(* IEC 61131-3 sources: volt/packages/volt-lsp-iec/test-corpus/lenze-mid/Device/Plc Logic/Application/Library Manager/AlarmManager, 462 files *)

(* ---- ACKNOWLEDGEMETHOD.dut ---- *)
TYPE ACKNOWLEDGEMETHOD :
(
	ACK := 1,
	REP := 2,
	REP_ACK := 3,
	ACK_REP := 6,
	ACK_REP_ACK := 7
);
END_TYPE

(* ---- ALARM_ID.dut ---- *)
TYPE ALARM_ID : UINT;
END_TYPE

(* ---- ALARMBASEPROPERTYINFO.dut ---- *)
TYPE ALARMBASEPROPERTYINFO :
STRUCT
	PVARADR : POINTER TO BYTE;
END_STRUCT
END_TYPE

(* ---- ALARMEVENT.dut ---- *)
TYPE ALARMEVENT :
STRUCT
	USIALARMGROUPID : ALARMGROUP_ID;
	UIALARMID : ALARM_ID;
	LIPUTINTOEVENTQUEUEAT : Timestamp;
END_STRUCT
END_TYPE

(* ---- ALARMGROUP_ID.dut ---- *)
TYPE ALARMGROUP_ID : USINT;
END_TYPE

(* ---- ALARMINDICES.dut ---- *)
TYPE ALARMINDICES :
STRUCT
	M_IALARMGROUPINDEX : INT;
	M_IALARMINDEX : INT;
	M_ICALLERINDEX : INT;
END_STRUCT
END_TYPE

(* ---- ALARMMANAGERCLIENTINFOSTRUCT.dut ---- *)
TYPE ALARMMANAGERCLIENTINFOSTRUCT :
STRUCT
	ITFALARMMANAGERCLIENT : IAlarmManagerClient;
	PARRITFRELEVANTALARMS : POINTER TO ARRAY [0..10] OF IAlarm;
	ICOUNTRELEVANTALARMSLOC : INT;
	DICOUNTRELEVANTALARMSREM : DINT;
	PARRITFACTIVEALARMS : POINTER TO ARRAY [0..10] OF IAlarm;
	ICOUNTACTIVEALARMS : INT;
	PARRITFALARMSFROMHISTORY : POINTER TO ARRAY [0..10] OF IAlarm2;
	PARRALARMSGRPFORHISTORY : POINTER TO ARRAY [0..10] OF POINTER TO AlarmGroupAdapter;
	PARRALARMSCLFORHISTORY : POINTER TO ARRAY [0..10] OF POINTER TO AlarmClassAdapter;
	ICOUNTALARMSFROMHISTORY : INT;
	PARRSTRUCTPROXYREGISTERED : POINTER TO ARRAY [0..10] OF StructProxyRegistered;
	IPROXYCNT : INT;
END_STRUCT
END_TYPE

(* ---- ALARMMANAGERGETALARMSEVENTPARAMS.dut ---- *)
TYPE ALARMMANAGERGETALARMSEVENTPARAMS :
STRUCT
	PSZAPPLNAME : POINTER TO STRING;
	ISKIPROWS : INT;
	IMAXROWS : INT;
	UDICOUNTALARMGROUPS : UDINT;
	PUIARRALARMGROUPS : POINTER TO ARRAY [0..0] OF UDINT;
	UDICOUNTALARMCLASSES : UDINT;
	PUIARRALARMCLASSES : POINTER TO ARRAY [0..0] OF UDINT;
	USIPRIORITYFROM : USINT;
	USIPRIORITYTO : USINT;
	BROWIDVALID : BOOL;
	DIROWID : DINT;
	PBRESULT : POINTER TO BYTE;
	UDIBUFFERSIZE : UDINT;
	UDICOUNTROWS : UDINT;
	UIERROR : UINT;
	BREQUESTHANDLED : BOOL;
END_STRUCT
END_TYPE

(* ---- ALARMMANAGERGETCOUNTEVENTPARAMS.dut ---- *)
TYPE ALARMMANAGERGETCOUNTEVENTPARAMS :
STRUCT
	PSZAPPLNAME : POINTER TO STRING;
	UDICOUNTALARMGROUPS : UDINT;
	PUIARRALARMGROUPS : POINTER TO ARRAY [0..0] OF UDINT;
	UDICOUNTALARMCLASSES : UDINT;
	PUIARRALARMCLASSES : POINTER TO ARRAY [0..0] OF UDINT;
	USIPRIORITYFROM : USINT;
	USIPRIORITYTO : USINT;
	UDICOUNT : UDINT;
	BREQUESTHANDLED : BOOL;
END_STRUCT
END_TYPE

(* ---- ALARMRECORD.dut ---- *)
TYPE ALARMRECORD :
STRUCT
	IRECORDID : INT := -1;
	UICLIENT : UINT;
	IALARMGROUP : INT;
	PAITFALARMGROUP : POINTER TO ARRAY [0..9] OF IAlarmGroup;
	IALARMCLASS : INT;
	PAITFALARMCLASS : POINTER TO ARRAY [0..9] OF IAlarmClass;
	IALARMCLASSINSERT : INT;
END_STRUCT
END_TYPE

(* ---- ALARMSTATE.dut ---- *)
TYPE ALARMSTATE :
(
	NOTDEFINED := 16#FF,
	NORMAL := 0,
	ACTIVE := 2,
	WAITINGFORCONFIRMATION := 3,
	ACTIVEACKNOWLEDGED := 4,
	INACTIVEUNACKNOWLEDGED := 5,
	PENDING := 1
);
END_TYPE

(* ---- ALARMSTATETRANSITION.dut ---- *)
TYPE ALARMSTATETRANSITION :
(
	NOTRANSITION := 0,
	PENDING := -1,
	ACTIVATE := 1,
	DEACTIVATE := 2,
	ACKNOWLEDGE := 3,
	CONFIRM := 4,
	REALARM := 5
);
END_TYPE

(* ---- ALARMSTORAGELATCHVARIABLE.dut ---- *)
TYPE ALARMSTORAGELATCHVARIABLE :
STRUCT
	M_BYTYPE : BYTE;
	M_LIVALUE : LINT;
	M_XVALUENULL : BOOL;
END_STRUCT
END_TYPE

(* ---- ALARMSTORAGESTATICDATA.dut ---- *)
TYPE ALARMSTORAGESTATICDATA :
STRUCT
	LITIMESTAPLAST : TIMESTAMP;
	LITIMESTAPACTIVE : TIMESTAMP;
	LITIMESTAPINACTIVE : TIMESTAMP;
	LITIMESTAPACKNOWLEDGE : TIMESTAMP;
	IOFFSETLAST : INT := -1;
	IOFFSETACTIVE : INT := -1;
	IOFFSETINACTIVE : INT := -1;
	IOFFSETACKNOWLEDGE : INT := -1;
	LITRIGGERVALUEVAL : LINT;
	ITRIGGERVALUETYPE : TypeClass;
	UDIALARMID : UDINT;
	UDIALARMGROUPID : UDINT;
	UDIALARMCLASSID : UDINT;
	ESTATE : AlarmState;
	USIPRIORITY : USINT;
	LIREMOTEDEVICEVAL : LINT;
	PWSCMTACTIVEACK : POINTER TO WSTRING;
	PWSCMTNORMAL : POINTER TO WSTRING;
	PWSCMTACTIVE : POINTER TO WSTRING;
	PWSCMTWAITINGCONF : POINTER TO WSTRING;
	PWSUSERIDACTIVEACK : POINTER TO WSTRING;
	PWSUSERIDNORMAL : POINTER TO WSTRING;
	PWSUSERIDACTIVE : POINTER TO WSTRING;
	PWSUSERIDWAITINGCONF : POINTER TO WSTRING;
	IDROW : CAA.IDENT;
END_STRUCT
END_TYPE

(* ---- ALARMSTRUCTFONT.dut ---- *)
TYPE ALARMSTRUCTFONT :
STRUCT
	SNAME : STRING := 'Arial';
	IHEIGHT : INT := 12;
	DWFLAGS : DWORD := 16#0;
	DWCHARSET : DWORD := 16#0;
	DWCOLOR : DWORD := 16#0;
END_STRUCT
END_TYPE

(* ---- ALARMUNIONBYTEORDERTEST.dut ---- *)
TYPE ALARMUNIONBYTEORDERTEST :
UNION
	W : WORD;
	BTS : ARRAY [0..1] OF BYTE;
END_UNION
END_TYPE

(* ---- CONFIGURABLEEXPRESSION.dut ---- *)
TYPE CONFIGURABLEEXPRESSION :
(
	OBSERVEDEXPRESSION := 0,
	LATCHVAR1 := 1,
	LATCHVAR2 := 2,
	LASTLATCHVARIABLE := 1000
);
END_TYPE

(* ---- DISPLAYOPTIONS.dut ---- *)
TYPE DISPLAYOPTIONS :
STRUCT
	FONT : AlarmStructFont;
	DWBACKGROUNDCOLOR : DWORD := 16#FFFFFF;
	SBITMAPID : STRING;
	XTRANSPARENT : BOOL;
	DWTRANSPARENTCOLOR : DWORD;
END_STRUCT
END_TYPE

(* ---- EALARMBYTEORDER.dut ---- *)
TYPE EALARMBYTEORDER :
(
	INTEL,
	MOTOROLA,
	UNKNOWN
);
END_TYPE

(* ---- EALARMCOMMENT.dut ---- *)
TYPE EALARMCOMMENT :
(
	NO_COMMENT,
	COMMENT_NORMAL,
	COMMENT_ACTIVE_ACK
);
END_TYPE

(* ---- EALARMCOMPARABLE.dut ---- *)
TYPE EALARMCOMPARABLE :
(
	FIRST_ENTRY := 0,
	TIMESTAMP_LAST := 0,
	TIMESTAMP_ACTIVE := 1,
	TIMESTAMP_INACTIVE := 2,
	TIMESTAMP_ACKNOWLEDGE := 3,
	VALUE := 4,
	MESSAGE := 5,
	PRIORITY := 6,
	ALARM_CLASS := 7,
	STATE := 8,
	REM_DEVICE := 9,
	COMMENT_ACK := 10,
	USERID_ACK := 11,
	LAST_ENTRY := 11
);
END_TYPE

(* ---- EALARMSTORAGEMIRRORSTATE.dut ---- *)
TYPE EALARMSTORAGEMIRRORSTATE :
(
	NOTYETMIRRORED,
	MIRRORINGSTARTED,
	ADDITIONALREADCALLREQUIRED,
	COMPLETELYMIRRORED,
	ERROR,
	RELOADREQUIRED
);
END_TYPE

(* ---- EALARMSTORAGEOBJECT.dut ---- *)
TYPE EALARMSTORAGEOBJECT :
(
	IX_MIN := 0,
	TBL_ALARM := IX_MIN,
	TBL_METADATA := 1,
	TBL_VERSION := 2,
	IDX_TSLAST := 3,
	IDX_GROUP_TSLAST := 4,
	IDX_CLASS_TSLAST := 5,
	TBL_LATCH_VAR_STRINGS := 6,
	IDX_LATCH_VAR_STRINGS := 7,
	IDX_LATCH1_TSLAST := 8,
	IX_LAST := IDX_LATCH1_TSLAST
);
END_TYPE

(* ---- EALARMSTORAGEREADERERRORS.dut ---- *)
TYPE EALARMSTORAGEREADERERRORS :
(
	NOERROR := CmpErrors.Errors.ERR_OK,
	WRONGPARAMETER := CmpErrors.Errors.ERR_PARAMETER,
	NOMEMORY := CmpErrors.Errors.ERR_NOMEMORY,
	NOOBJECT := CmpErrors.Errors.ERR_NO_OBJECT,
	ADDITIONALREADCALLREQUIRED := CmpErrors.Errors.ERR_PENDING,
	INVALIDCALL := 20002
);
END_TYPE

(* ---- EALARMTYPE.dut ---- *)
TYPE EALARMTYPE :
(
	UNDEFINED := 0,
	ALARM := 1,
	EVENT := 2,
	IMPLICITLYACKNOWLEDGEDEVENT := 3,
	ALARMAPI := 4
);
END_TYPE

(* ---- ECOMPARABLETYPE.dut ---- *)
TYPE ECOMPARABLETYPE :
(
	TYPE_UNDEFINED := 0,
	TYPE_BOOL := 1,
	TYPE_NUMERIC := 2,
	TYPE_STRING := 3
);
END_TYPE

(* ---- EDBACTIVEINDEX.dut ---- *)
TYPE EDBACTIVEINDEX :
(
	NOT_DEFINED := 0,
	TIMESTAMP,
	GROUP,
	EDB_CLASS,
	LATCH1
);
END_TYPE

(* ---- EDBTYPE.dut ---- *)
TYPE EDBTYPE :
(
	NOT_DEFINED := 0,
	SQL,
	MEMORY
);
END_TYPE

(* ---- EFILTERLATCHCONTENT.dut ---- *)
TYPE EFILTERLATCHCONTENT :
(
	NOT_SET := -1,
	DISABLE := 0,
	STR := 1,
	IEC := 2,
	NUMBER := 3
);
END_TYPE

(* ---- EFILTERTIMERANGETYPE.dut ---- *)
TYPE EFILTERTIMERANGETYPE :
(
	NOT_SET := -1,
	DISABLE := 0,
	ENABLE := 1
);
END_TYPE

(* ---- ELOCALBUFFERCURSORSTATE.dut ---- *)
TYPE ELOCALBUFFERCURSORSTATE :
(
	EOF := -3,
	CLOSED := -2,
	OPEN := -1
);
END_TYPE

(* ---- ENUMERICCOMPARISON.dut ---- *)
TYPE ENUMERICCOMPARISON :
(
	AS_LINT := 0,
	AS_REAL := 1,
	AS_LREAL := 2
);
END_TYPE

(* ---- EVTPARAM_CHANNELCLOSED.dut ---- *)
TYPE EVTPARAM_CHANNELCLOSED :
STRUCT
	UICLIENT : UINT;
	UICHANNELHANDLE : UINT;
	ERRREASON : RTS_IEC_RESULT;
END_STRUCT
END_TYPE

(* ---- FILELIMIT.dut ---- *)
TYPE FILELIMIT :
(
	NOLIMIT := 0,
	RECORDS := 1,
	SIZE := 2
);
END_TYPE

(* ---- HISTORICALACTIVEALARMROWID.dut ---- *)
TYPE HISTORICALACTIVEALARMROWID :
STRUCT
	DWROWID : DWORD;
	LITS : LINT;
END_STRUCT
END_TYPE

(* ---- LATCHVARIABLE.dut ---- *)
TYPE LATCHVARIABLE :
STRUCT
	M_BYTYPE : BYTE;
	M_LIVALUE : LINT;
END_STRUCT
END_TYPE

(* ---- LOCALBUFFERDATABASEACCESSCONTEXT.dut ---- *)
TYPE LOCALBUFFERDATABASEACCESSCONTEXT :
STRUCT
	M_HSEMTRANSACTION : RTS_IEC_HANDLE := RTS_INVALID_HANDLE;
	M_DICURSORINDEX : DINT := ELocalBufferCursorState.Closed;
	M_PALICURRALARM : POINTER TO ARRAY [0..0] OF LINT;
	M_CBPSTRINGLATCHVARIABLE : CharBufferPtr;
	M_XISONLYONEALARMGROUPSELECTED : BOOL;
	M_XISONLYONEALARMCLASSSELECTED : BOOL;
	M_ELASTERROR : STO.ERROR;
END_STRUCT
END_TYPE

(* ---- MONITORDBSTATUS.dut ---- *)
TYPE MONITORDBSTATUS :
STRUCT
	DBTYPE : EDBType;
	ACTIVEINDEX : EDBActiveIndex;
	IERROR : INT;
	SFUNCTION : STRING;
	IACTION : INT;
END_STRUCT
END_TYPE

(* ---- MONITORFILTERBYDATETIME.dut ---- *)
TYPE MONITORFILTERBYDATETIME :
STRUCT
	FILTERTARGET : EFilterTimeRangeType;
	DTFROMVALUE : DATE_AND_TIME;
	DTTOVALUE : DATE_AND_TIME;
END_STRUCT
END_TYPE

(* ---- MONITORFILTERBYLATCH.dut ---- *)
TYPE MONITORFILTERBYLATCH :
STRUCT
	FILTERLATCHCONTENT : EFilterLatchContent;
	VTYPE : Visu_Types;
	LIVALUE : LINT;
	RVALUE : REAL;
	LRVALUE : LREAL;
	WSSTRVALUE : WSTRING(255);
END_STRUCT
END_TYPE

(* ---- PLACEHOLDERANALYZATIONSTATE.dut ---- *)
TYPE PLACEHOLDERANALYZATIONSTATE :
(
	NOTAVAILABLE := 16#0,
	TOOMANYPLACEHOLDERS := 16#1,
	INVALIDPLACEHOLDER := 16#2,
	CYCLICALLYREPAINTREQUIRED := 16#4,
	DONE := 16#10
);
END_TYPE

(* ---- PLACEHOLDERDESCRIPTION.dut ---- *)
TYPE PLACEHOLDERDESCRIPTION :
STRUCT
	M_EPLACEHOLDER : Placeholder;
	M_PCBSPLACEHOLDER : POINTER TO CharBufferString;
	M_XSUPPORTSFORMATSTRING : BOOL;
	M_XINHIBITSOPTIMIZATION : BOOL;
	M_XREQUIREDCYCLICALLYREPAINT : BOOL;
	M_XINHIBITMULTIPLEUSAGE : BOOL;
	M_PCBSRELATEDPLACEHOLDERSUBSTRING : POINTER TO CharBufferString;
	M_PCBSRELATEDPLACEHOLDERBRACKET : POINTER TO CharBufferString;
END_STRUCT
END_TYPE

(* ---- PLACEHOLDERINFO.dut ---- *)
TYPE PLACEHOLDERINFO :
STRUCT
	M_APLACEHOLDEROCCURRENCE : ARRAY [0..(AlarmConstants.COUNT_PLACEHOLDER - 1)] OF PlaceholderOccurrence;
	M_SICOUNTPLACEHOLDERS : SINT := -1;
	M_EPLACEHOLDERANALYZATIONSTATE : PlaceholderAnalyzationState;
END_STRUCT
END_TYPE

(* ---- PLACEHOLDERSCANNERSTATE.dut ---- *)
TYPE PLACEHOLDERSCANNERSTATE :
(
	START := 0,
	SKIPWHITESPACE := 1,
	SCANFORMAT := 2,
	END := 3,
	ERROR := 255
);
END_TYPE

(* ---- PROXYENUMSTATE.dut ---- *)
TYPE PROXYENUMSTATE :
(
	NOTRUNNING,
	PREPARATION,
	CHECKDATA,
	RUN
);
END_TYPE

(* ---- PROXYSTRUCTALARM.dut ---- *)
TYPE PROXYSTRUCTALARM :
STRUCT
	UIALARMID : ALARM_ID;
	UDIALARMINTERNALID : UDINT;
	UDIALARMGROUPINTERNALID : UDINT;
	UDIALARMCLASSINTERNALID : UDINT;
	SALARMID : STRING;
	XACK : BOOL;
END_STRUCT
END_TYPE

(* ---- PROXYSTRUCTALARMCLASS.dut ---- *)
TYPE PROXYSTRUCTALARMCLASS :
STRUCT
	UDIINTERNALID : UDINT;
	SNAME : STRING;
	USIPRIORITY : USINT;
	XACKNOWLEDGESEPARATELY : BOOL;
	ADISPLAYOPTIONS : ARRAY [AlarmState.Normal..AlarmState.ActiveAcknowledged] OF DisplayOptions;
	AXDISPLAYOPTIONSSET : ARRAY [AlarmState.Normal..AlarmState.ActiveAcknowledged] OF BOOL;
END_STRUCT
END_TYPE

(* ---- PROXYSTRUCTALARMCLASSDESC.dut ---- *)
TYPE PROXYSTRUCTALARMCLASSDESC :
STRUCT
	XVALID : BOOL;
	SNAME : STRING;
	USIPRIORITY : USINT;
	UDIINTERNALID : UDINT;
END_STRUCT
END_TYPE

(* ---- PROXYSTRUCTALARMDESC.dut ---- *)
TYPE PROXYSTRUCTALARMDESC :
STRUCT
	XVALID : BOOL;
	SALARMID : STRING;
	UIALARMID : ALARM_ID;
	UDIALARMINTERNALID : UDINT;
	UDIALARMGROUPINTERNALID : UDINT;
END_STRUCT
END_TYPE

(* ---- PROXYSTRUCTALARMGROUP.dut ---- *)
TYPE PROXYSTRUCTALARMGROUP :
STRUCT
	UDIINTERNALID : UDINT;
	SNAME : STRING;
	STEXTLIST : STRING;
END_STRUCT
END_TYPE

(* ---- PROXYSTRUCTALARMGROUPDESC.dut ---- *)
TYPE PROXYSTRUCTALARMGROUPDESC :
STRUCT
	XVALID : BOOL;
	SNAME : STRING;
	STEXTLIST : STRING;
	UDIINTERNALID : UDINT;
END_STRUCT
END_TYPE

(* ---- PROXYSTRUCTCLASSREMAP.dut ---- *)
TYPE PROXYSTRUCTCLASSREMAP :
STRUCT
	SCLASSORIGINAL : STRING;
	SCLASSNEW : STRING;
END_STRUCT
END_TYPE

(* ---- PROXYSTRUCTDSCHANNELPARAM.dut ---- *)
TYPE PROXYSTRUCTDSCHANNELPARAM :
STRUCT
	ITFDATASOURCESMGR : IDatasources.IDatasourcesMgr;
	PSDSNAME : POINTER TO STRING;
	ILATCHVARSNUM : INT;
	PSALMSTATETRANSCOUNTER : POINTER TO STRING;
	PALMSTATETRANSCOUNTER : __XWORD;
	TYPEALMSTATETRANSCOUNTER : TypeClass;
	PSALMSTORAGECOUNTER : POINTER TO STRING;
	PALMSTORAGECOUNTER : __XWORD;
	TYPEALMSTORAGECOUNTER : TypeClass;
END_STRUCT
END_TYPE

(* ---- PROXYSTRUCTERROR.dut ---- *)
TYPE PROXYSTRUCTERROR :
STRUCT
	UDIERROR : UDINT;
	LTTIMESTAMP : LTIME;
	SMSG : STRING(20);
END_STRUCT
END_TYPE

(* ---- PROXYSTRUCTHISTORICALALARMACTIVE.dut ---- *)
TYPE PROXYSTRUCTHISTORICALALARMACTIVE :
STRUCT
	DWROWIDLOCAL : DWORD := AlarmConstants.INVALID_ROWID;
	DWROWIDREMOTE : DWORD := AlarmConstants.INVALID_ROWID;
	LITSACTIVEREMOTE : LINT;
	ESTATELAST : AlarmState := AlarmState.NotDefined;
END_STRUCT
END_TYPE

(* ---- PROXYSTRUCTINITIALIZE.dut ---- *)
TYPE PROXYSTRUCTINITIALIZE :
STRUCT
	PSPROXYNAME : POINTER TO STRING;
	ITFPROXYCOMMCHANNEL : IProxyCommChannel;
	PSAPPNAME : POINTER TO STRING;
	PAALARMGROUPS : POINTER TO ARRAY [0..9] OF STRING;
	IALARMGROUPSNUM : INT;
	PACLASSREMAP : POINTER TO ARRAY [0..9] OF ProxyStructClassReMap;
	ICLASSREMAPNUM : INT;
END_STRUCT
END_TYPE

(* ---- PROXYSTRUCTMONITOR.dut ---- *)
TYPE PROXYSTRUCTMONITOR :
STRUCT
	SNAME : STRING;
	ESTATE : ProxyEnumState;
	IALARMCLASSNUM : INT;
	IALARMGROUPSNUM : INT;
	DIALARMNUM : DINT;
	ILATCHVARSNUM : INT;
	IACTIVEALARMS : INT;
	DIHISTACTIVEALMSCNT : DINT;
	IHISTROWALMSCNT : INT;
	IHISTROWACTIVEALMSCNT : INT;
	XHASSTORAGE : BOOL;
	DWROWIDFIRSTREMDB : DWORD;
	DWROWIDLASTREMDB : DWORD;
	DWROWIDLASTLOCDB : DWORD;
	DIWRITEDBCNTTOT : DINT;
	IWRITEDBCNT : INT;
	TWRITEDBDURATIONLAST : TIME;
	DITOTMEM : DINT;
	DIHISTACTIVEALMSSIZE : DINT;
	IHISTROWALMSSIZE : INT;
	IHISTROWACTIVEALMSSIZE : INT;
	LIBVERALMMAN : VERSION;
END_STRUCT
END_TYPE

(* ---- PROXYSTRUCTMONITORALARMCLASSDESC.dut ---- *)
TYPE PROXYSTRUCTMONITORALARMCLASSDESC :
STRUCT
	SNAME : STRING;
	UDIINTERNALID : UDINT;
	USIPRIORITY : USINT;
	XACKNOWLEDGESEPARATELY : BOOL;
END_STRUCT
END_TYPE

(* ---- PROXYSTRUCTMONITORALARMDESC.dut ---- *)
TYPE PROXYSTRUCTMONITORALARMDESC :
STRUCT
	SALARMID : STRING;
	UIALARMID : ALARM_ID;
	UDIALARMINTERNALID : UDINT;
	UDIALARMGROUPINTERNALID : UDINT;
	UDIALARMCLASSINTERNALID : UDINT;
END_STRUCT
END_TYPE

(* ---- PROXYSTRUCTMONITORALARMGROUPDESC.dut ---- *)
TYPE PROXYSTRUCTMONITORALARMGROUPDESC :
STRUCT
	SNAME : STRING;
	UDIINTERNALID : UDINT;
	STEXTLIST : STRING;
END_STRUCT
END_TYPE

(* ---- PROXYSTRUCTMONITORREQUEST.dut ---- *)
TYPE PROXYSTRUCTMONITORREQUEST :
STRUCT
	ITASKID : INT := ProxyConstants.REQ_ID_NONE;
	AFIFOERRORS : ARRAY [1..ProxyConstants.FIFO_ERROR_SIZE] OF ProxyStructError;
	UDIERRCOUNT : UDINT;
	LTELAPTIME : LTIME;
	TREQDURATIONLAST : TIME;
	TREQDURATIONAVG : TIME;
	TREQDURATIONMIN : TIME;
	TREQDURATIONMAX : TIME;
	UDIREQDURATIONBUILDREQ : UDINT;
	UDIREQDURATIONWAITANS : UDINT;
	UDIREQDURATIONELABANS : UDINT;
	UDIREQCOUNT : UDINT;
	UDIREQCOUNTCLOSED : UDINT;
END_STRUCT
END_TYPE

(* ---- PROXYSTRUCTPARAM.dut ---- *)
TYPE PROXYSTRUCTPARAM :
STRUCT
	DWBASETIME : DWORD;
	DWACTALMTIME : DWORD;
	DWHISALMTIME : DWORD;
	DWACKALMTIME : DWORD;
	TTIMEOUT : TIME := TIME#5s0ms;
END_STRUCT
END_TYPE

(* ---- PROXYSTRUCTRECORD.dut ---- *)
TYPE PROXYSTRUCTRECORD :
STRUCT
	IRECORDID : INT;
	IALARMCLASSNUM : INT;
	DIALARMNUM : DINT;
	ILATCHVARSNUM : INT;
	PAALARMGROUPS : POINTER TO ARRAY [0..9] OF STRING;
	IALARMGROUPSNUM : INT;
	PACLASSREMAP : POINTER TO ARRAY [0..9] OF ProxyStructClassReMap;
	ICLASSREMAPNUM : INT;
	PAACTIVEALARMOBJSTUBS : POINTER TO ARRAY [0..100] OF POINTER TO ProxyFbAlarmMetaObjectStub;
	DIALMOBJSTUBSALLOC : DINT;
	PAACTIVEALARMCONTAINER : POINTER TO ARRAY [0..100] OF POINTER TO AlarmContainer;
	DIALMCONTAINERALLOC : DINT;
	DIACTIVEALARMS : DINT;
	PASTRUCTALARMDESCRIPTION : POINTER TO ARRAY [0..100] OF POINTER TO ProxyStructAlarm;
	DIALARMDESCALLOC : DINT;
	PASTRUCTALARMGROUPDESCRIPTION : POINTER TO ARRAY [0..100] OF POINTER TO ProxyStructAlarmGroup;
	IALARMGROUPDESCALLOC : INT;
	PASTRUCTALARMCLASSDESCRIPTION : POINTER TO ARRAY [0..100] OF POINTER TO ProxyStructAlarmClass;
	IALARMCLASSDESCALLOC : INT;
END_STRUCT
END_TYPE

(* ---- PROXYSTRUCTTASKCALL.dut ---- *)
TYPE PROXYSTRUCTTASKCALL :
STRUCT
	ITASKID : INT;
	DWSCHEDUL : DWORD;
	TTIMEOUT : TIME;
	XDONEOK : BOOL;
	XLOCK : BOOL;
	HLOCK : RTS_IEC_HANDLE;
	DWSCHEDULCNT : DWORD;
END_STRUCT
END_TYPE

(* ---- SCALARTYPE.dut ---- *)
TYPE SCALARTYPE :
UNION
	COMPBYTE : BYTE;
	COMPWORD : WORD;
	COMPDWORD : DWORD;
	COMPLWORD : LWORD;
	COMPSINT : SINT;
	COMPUSINT : USINT;
	COMPINT : INT;
	COMPUINT : UINT;
	COMPDINT : DINT;
	COMPUDINT : UDINT;
	COMPLINT : LINT;
	COMPULINT : ULINT;
	COMPBOOL : BOOL;
	COMPREAL : REAL;
	COMPLREAL : LREAL;
END_UNION
END_TYPE

(* ---- SQLITEDATABASEACCESSCONTEXT.dut ---- *)
TYPE SQLITEDATABASEACCESSCONTEXT :
STRUCT
	M_ITFTABLELATCHVARVALUES : STO.ITable;
	M_ITFCURSORLATCHVARVALUES : STO.ICursor;
	M_ITFROWLATCHVARVALUES : STO.IRow;
	M_IDTBLLATCHVARSTRINGS : CAA.IDENT;
	M_IDIDXLATCHVARSTRINGS : CAA.IDENT;
	M_ITFTRANSACTION : STO.ITransaction;
	M_ITFTABLE : STO.ITable;
	M_ITFCURSOR : STO.ICursor;
	M_ITFROW : STO.IRow;
	M_IDINDEX : CAA.IDENT;
	M_EINDEX : EAlarmStorageObject;
	M_ELASTERROR : STO.ERROR;
END_STRUCT
END_TYPE

(* ---- STORAGETASKINFO.dut ---- *)
TYPE STORAGETASKINFO :
STRUCT
	XTASKACTIVE : BOOL;
	PTASKINFO : POINTER TO CmpIecTask.Task_Info2;
END_STRUCT
END_TYPE

(* ---- STRINGCONTAINERBUFFERINFO.dut ---- *)
TYPE STRINGCONTAINERBUFFERINFO :
STRUCT
	PUDIBUFFERSIZE : POINTER TO UDINT;
	PUDIFIRSTFREEPOSITION : POINTER TO UDINT;
	PBYFIRSTPOSITION : POINTER TO BYTE;
	PBYFIRSTFREEPOSITION : POINTER TO BYTE;
END_STRUCT
END_TYPE

(* ---- STRUCTPROXYREGISTERED.dut ---- *)
TYPE STRUCTPROXYREGISTERED :
STRUCT
	ITFPROXY : IProxy;
	DIALM : DINT;
END_STRUCT
END_TYPE

(* ---- STRUFILTERREMOTEALM.dut ---- *)
TYPE STRUFILTERREMOTEALM :
STRUCT
	SPROXYNAME : STRING;
	DIID : DINT;
END_STRUCT
END_TYPE

(* ---- SWAPHELPER_UNION.dut ---- *)
TYPE SWAPHELPER_UNION :
UNION
	COMPBYTE : BYTE;
	COMPWORD : WORD;
	COMPDWORD : DWORD;
	COMPLWORD : LWORD;
END_UNION
END_TYPE

(* ---- TIMESTAMP.dut ---- *)
TYPE TIMESTAMP : LINT;
END_TYPE

(* ---- ALARMCONSTANTS.gvl ---- *)
VAR_GLOBAL
	NULL : POINTER TO BYTE := 0;
	MAX_PLACEHOLDER_LENGTH : BYTE := 25;
	MAX_PLACEHOLDER_REPLACEMENT_LENGTH : WORD := 255;
	REPL_AMP_ANSI : DWORD := 16#0;
	REPL_AMP_UNICODE : DWORD := 16#1;
	ALARM_MESSAGEBUFFER_SIZE : WORD := 500;
	MAX_MESSAGE_SIZE : WORD := 256;
	ALARM_SEPARATOR : STRING(1) := '$T';
	ALARMGROUP_SEPARATOR : STRING(1) := '|';
	SLEEP_TIME : UDINT := 5;
	RETRY_COUNT : INT := 10;
	NOT_RELEVANT : ALARM_ID := 65535;
	TICKS_1_1_1970 : ULINT := 116444736000000000;
	DIVISOR_TO_SECONDS : LINT := ((1000 * 1000) * 10);
	FMT_INT : BYTE := 0;
	FMT_LONG : BYTE := 1;
	FMT_FLOAT : BYTE := 2;
	FMT_STRING : BYTE := 3;
	FMT_WSTRING : BYTE := 4;
	FMT_FIRST_FORMAT_STRING : BYTE := FMT_INT;
	FMT_LAST_FORMAT_STRING : BYTE := FMT_WSTRING;
	PLH_FIRST_PLACEHOLDER : Placeholder := Placeholder.PLH_ALARM;
	PLH_LAST_PLACEHOLDER : Placeholder := Placeholder.PLH_TRIGGERVALUE;
	COUNT_PLACEHOLDER : BYTE := 22;
	INVALID_ROWID : CAA.IDENT := 0;
	LESS : INT := -1;
	EQUAL : INT := 0;
	GREATER : INT := 1;
	RECORD_ID_TEST : INT := 16#7FFF;
	RECORD_ID_TEST2 : INT := 16#7FFE;
	MAX_LATCH_VARS : INT := 10;
	SIZE_HIST_ACTIVE_ALM : INT := 250;
	VISU_TYPES_TYPE_LDATE : INT := 33;
	VISU_TYPES_TYPE_LDT : INT := 34;
	VISU_TYPES_TYPE_LTOD : INT := 35;
	ALARM_STORAGE_TASK_NAME : STRING := 'Visu_AlarmStorageTask';
END_VAR

(* ---- ALARMGLOBALS.gvl ---- *)
VAR_GLOBAL
	G_ACK_ALARMSTATEMACHINE : Ack_AlarmStateMachine;
	G_ACK_REP_ALARMSTATEMACHINE : Ack_Rep_AlarmStateMachine;
	G_ACK_REP_ACK_ALARMSTATEMACHINE : Ack_Rep_Ack_AlarmStateMachine;
	G_REP_ACK_ALARMSTATEMACHINE : Rep_Ack_AlarmStateMachine;
	G_REP_ALARMSTATEMACHINE : Rep_AlarmStateMachine;
	G_ACK_ALARMSTATEMACHINE_NOCONFIRM : Ack_AlarmStateMachine_NoConfirm;
	G_ACK_REP_ALARMSTATEMACHINE_NOCONFIRM : Ack_Rep_AlarmStateMachine_NoConfirm;
	G_ACK_REP_ACK_ALARMSTATEMACHINE_NOCONFIRM : Ack_Rep_Ack_AlarmStateMachine_NoConfirm;
	G_REP_ACK_ALARMSTATEMACHINE_NOCONFIRM : Rep_Ack_AlarmStateMachine_NoConfirm;
	G_ALARMHANDLER_INST : StandardAlarmHandler;
	G_ALARMHANDLER : IAlarmHandler9 := g_AlarmHandler_Inst;
	G_ALARMHANDLERBASE : IAlarmHandlerBase := g_AlarmHandler_Inst;
	G_ALARMHANDLERREMOTE : IAlarmHandlerRemote := g_AlarmHandler_Inst;
	G_ALARMHANDLERREMOTEMONITOR : IAlarmHandlerRemoteMonitor := g_AlarmHandler_Inst;
	G_ALARMSTORAGEQUEUE : AlarmStorageQueue;
	G_DIALARMSTATETRANSITIONCOUNTER : DINT;
	G_DIALARMSTORAGECOUNTER : DINT;
	STATE : INT;
	G_STAPPLICATIONNAME : STRING;
	G_PAPPLICATION : POINTER TO CmpApp.APPLICATION := RTS_INVALID_HANDLE;
	G_ERRORHANDLER : DatabaseAccessErrorHandler;
	G_BBYTEORDERDETERMINED : BOOL := FALSE;
	G_XMETADATAFILECREATED : BOOL := FALSE;
	G_SDATEFORMAT : STRING := 'dd.MM.yyyy';
	G_STIMEFORMAT : STRING := 'HH:mm:ss';
	G_DATEFORMATTER : STU.DateFormatter;
	G_TIMEFORMATTER : STU.TimeFormatter;
	G_TYPEDVALUEFORMATTER : TypedValueFormatter;
	G_SALARMSTATETEXTLISTNAME : STRING := 'AlarmManager.TL_AlarmStatus';
	COMPONENT_NAME : STRING := 'AlarmManager';
	G_STRINGPLACEHOLDERDATE : CharBufferString;
	G_STRINGPLACEHOLDERDATE2 : CharBufferString;
	G_STRINGPLACEHOLDERALLDEFAULT : CharBufferString;
	G_STRINGPLACEHOLDERMESSAGE : CharBufferString;
	G_STRINGPLACEHOLDERTIME : CharBufferString;
	G_STRINGPLACEHOLDERTIME2 : CharBufferString;
	G_STRINGPLACEHOLDERSTATE : CharBufferString;
	G_STRINGPLACEHOLDERSTATE2 : CharBufferString;
	G_STRINGPLACEHOLDEREXPRESSION : CharBufferString;
	G_STRINGPLACEHOLDEREXPRESSION2 : CharBufferString;
	G_STRINGPLACEHOLDERPRIORITY : CharBufferString;
	G_STRINGPLACEHOLDERPRIORITY2 : CharBufferString;
	G_STRINGPLACEHOLDERCLASS : CharBufferString;
	G_STRINGPLACEHOLDERCLASS2 : CharBufferString;
	G_STRINGPLACEHOLDERALARMID : CharBufferString;
	G_STRINGPLACEHOLDERCURRENTVALUE : CharBufferString;
	G_STRINGPLACEHOLDERCURRENTVALUE2 : CharBufferString;
	G_STRINGPLACEHOLDERTRIGGERVALUE : CharBufferString;
	G_STRINGPLACEHOLDERTRIGGERVALUE2 : CharBufferString;
	G_STRINGPLACEHOLDERLATCH : CharBufferString;
	G_STRINGPLACEHOLDERLATCHWITHOPENINGBRACKET : CharBufferString;
	G_STRINGPLACEHOLDERALARM : CharBufferString;
	G_WSTRINGPLACEHOLDERDATE : CharBufferString;
	G_WSTRINGPLACEHOLDERDATE2 : CharBufferString;
	G_WSTRINGPLACEHOLDERALLDEFAULT : CharBufferString;
	G_WSTRINGPLACEHOLDERMESSAGE : CharBufferString;
	G_WSTRINGPLACEHOLDERTIME : CharBufferString;
	G_WSTRINGPLACEHOLDERTIME2 : CharBufferString;
	G_WSTRINGPLACEHOLDERSTATE : CharBufferString;
	G_WSTRINGPLACEHOLDERSTATE2 : CharBufferString;
	G_WSTRINGPLACEHOLDEREXPRESSION : CharBufferString;
	G_WSTRINGPLACEHOLDEREXPRESSION2 : CharBufferString;
	G_WSTRINGPLACEHOLDERPRIORITY : CharBufferString;
	G_WSTRINGPLACEHOLDERPRIORITY2 : CharBufferString;
	G_WSTRINGPLACEHOLDERCLASS : CharBufferString;
	G_WSTRINGPLACEHOLDERCLASS2 : CharBufferString;
	G_WSTRINGPLACEHOLDERALARMID : CharBufferString;
	G_WSTRINGPLACEHOLDERCURRENTVALUE : CharBufferString;
	G_WSTRINGPLACEHOLDERCURRENTVALUE2 : CharBufferString;
	G_WSTRINGPLACEHOLDERTRIGGERVALUE : CharBufferString;
	G_WSTRINGPLACEHOLDERTRIGGERVALUE2 : CharBufferString;
	G_WSTRINGPLACEHOLDERLATCH : CharBufferString;
	G_WSTRINGPLACEHOLDERLATCHWITHOPENINGBRACKET : CharBufferString;
	G_WSTRINGPLACEHOLDERALARM : CharBufferString;
	G_APSTRINGPLACEHOLDERS : ARRAY [AlarmConstants.PLH_FIRST_PLACEHOLDER..AlarmConstants.PLH_LAST_PLACEHOLDER] OF POINTER TO CharBufferString;
	G_APWSTRINGPLACEHOLDERS : ARRAY [AlarmConstants.PLH_FIRST_PLACEHOLDER..AlarmConstants.PLH_LAST_PLACEHOLDER] OF POINTER TO CharBufferString;
	G_APSTRINGPLACEHOLDERSBRACKET : ARRAY [AlarmConstants.PLH_FIRST_PLACEHOLDER..AlarmConstants.PLH_LAST_PLACEHOLDER] OF POINTER TO CharBufferString;
	G_APWSTRINGPLACEHOLDERSBRACKET : ARRAY [AlarmConstants.PLH_FIRST_PLACEHOLDER..AlarmConstants.PLH_LAST_PLACEHOLDER] OF POINTER TO CharBufferString;
	G_DATETIMEPLACEHOLDER : OnlyDateAndTimePlaceholder;
	G_EMPTYLATCHVARIABLE : ValueTypeBundle;
	G_RUNTIMEEVENTLISTENER : RuntimeEventListener;
	G_ALARMSTATECHANGEDEVENTLISTENER : AlarmStateChangedEventListener;
	G_STRINGCONTAINER : StringContainer;
	G_AWTEMPBUFFER : ARRAY [0..255] OF WORD;
	G_IPROXYQUEUESIZEHISTORICALALARM : INT := 300;
	G_IPROXYQUEUESIZEACTIVEHISTORICALALARM : INT := 100;
	G_XPLACEHOLDERREPLACEMENTFORMESSAGESORTING : BOOL := FALSE;
	G_IALARMSTORAGECLEAR : INT;
	G_ALARMLOCALSTORAGELIMIT : AlarmStorageLimit;
	G_IPERCDBALARMLIMIT : INT := 5;
	G_RRECORDSIZEFACTOR : REAL := 2.5;
	G_ITESTFAILREORD : INT;
	G_BDENYDATABASETRANSACTION : BOOL := FALSE;
	G_STORAGETASK_INST : CmpIecTask.Task_Info2;
	G_STORAGETASKINFO : StorageTaskInfo;
	G_ALARMALLOC : Allocator;
	G_INITALARMSONSTARTUP : VisuShared.Visu_FbInitOnStartup;
	G_BFIRSTCYCLEAFTERONLINECHANGE : BOOL;
	G_BFIRSTCYCLEAFTERDOWNLOAD : BOOL := TRUE;
	G_BALARMSDISABLED : BOOL;
	G_XSTEPBYSTEPMODE : BOOL := TRUE;
	G_TSTEPBYSTEPLIMIT : TIME := TIME#25ms;
END_VAR

(* ---- ALARMMANAGERBENCHMARKS.gvl ---- *)
VAR_GLOBAL
	ALARMSTORAGESTATISTICS : AlarmManagerRealValueStatistics;
END_VAR

(* ---- ALARMONLINECHANGEGLOBALS.gvl ---- *)
VAR_GLOBAL
	G_ACTIVEALARMSSTORAGE : ActiveAlarmsTempStorage;
END_VAR

(* ---- ALARMPARAMS.gvl ---- *)
VAR_GLOBAL
	PLACEHOLDER_VALUE_LENGTH : INT := (ANY_TO_INT(60) * ANY_TO_INT(2));
	COUNT_ROWS_TO_CHECK_FOR_OLDEST_ALARMS : INT := 50;
END_VAR

(* ---- ALARMSTORAGEREADERGLOBALS.gvl ---- *)
VAR_GLOBAL
	G_IMAXCOUNTROWSTOREAD : INT := 1000;
END_VAR

(* ---- ALARMSYNCGLOBALS.gvl ---- *)
VAR_GLOBAL
	HLOCKACTIVEALARMS : RTS_IEC_HANDLE := RTS_INVALID_HANDLE;
	HLOCKALLALARMS : RTS_IEC_HANDLE := RTS_INVALID_HANDLE;
	HLOCKALARMSTORAGEQUEUE : RTS_IEC_HANDLE := RTS_INVALID_HANDLE;
	BALARMSTORAGEINITIALIZED : BOOL := FALSE;
	BALARMSTORAGETASKACTIVE : BOOL := FALSE;
END_VAR

(* ---- ALARMTESTCONSTANTS.gvl ---- *)
VAR_GLOBAL
	G_TESTTIMESTAMPS : ARRAY [0..60] OF ULINT := [1706255000000, 1706255050000, 1706255100000, 1706255150000, 1706255200000, 1706255250000, 1706255300000, 1706255350000, 1706255400000, 1706255450000, 1706255500000, 1706255550000, 1706255600000, 1706255650000, 1706255700000, 1706255750000, 1706255800000, 1706255850000, 1706255900000, 1706255950000, 1706256000000, 1706256050000, 1706256100000, 1706256150000, 1706256200000, 1706256250000, 1706256300000, 1706256350000, 1706256400000, 1706256450000, 1706256500000, 1706256550000, 1706256600000, 1706256650000, 1706256700000, 1706256750000, 1706256800000, 1706256850000, 1706256900000, 1706256950000, 1706257000000, 1706257050000, 1706257100000, 1706257150000, 1706257200000, 1706257250000, 1706257300000, 1706257350000, 1706257400000, 1706257450000, 1706257500000, 1706257550000, 1706257600000, 1706257650000, 1706257700000, 1706257750000, 1706257800000, 1706257850000, 1706257900000, 1706257950000, 1706258000000];
	G_ICURRENTUSEDTIMESTAMP : INT := 0;
END_VAR

(* ---- ALARMTESTING.gvl ---- *)
VAR_GLOBAL
	XBLOCKSTORAGE : BOOL;
	XSTOREALARMS : BOOL;
	XRESTOREALARMS : BOOL;
	COMPILECHECKONLY : BOOL;
END_VAR

(* ---- ALARMVERSIONCONSTANTS.gvl ---- *)
VAR_GLOBAL
	_ALARMMANAGER_VERSION_LARGEROREQUAL_3_5_1_0_ : INT := 0;
	_ALARMMANAGER_VERSION_LARGEROREQUAL_3_5_3_40_ : INT := 0;
	_ALARMMANAGER_VERSION_LARGEROREQUAL_3_5_6_0_ : INT := 0;
	_ALARMMANAGER_VERSION_LARGEROREQUAL_3_5_7_0_ : INT := 0;
	_ALARMMANAGER_VERSION_LARGEROREQUAL_3_5_8_0_ : INT := 0;
	_ALARMMANAGER_VERSION_LARGEROREQUAL_3_5_9_0_ : INT := 0;
	_ALARMMANAGER_VERSION_LARGEROREQUAL_3_5_9_50_ : INT := 0;
	_ALARMMANAGER_VERSION_LARGEROREQUAL_3_5_10_0_ : INT := 0;
	_ALARMMANAGER_VERSION_LARGEROREQUAL_3_5_12_0_ : INT := 0;
	_ALARMMANAGER_VERSION_LARGEROREQUAL_3_5_13_0_ : INT := 0;
	_ALARMMANAGER_VERSION_LARGEROREQUAL_3_5_15_0_ : INT := 0;
	_ALARMMANAGER_VERSION_LARGEROREQUAL_3_5_16_0_ : INT := 0;
END_VAR

(* ---- COMPONENTCONSTANTS.gvl ---- *)
VAR_GLOBAL
	COMPONENTNAME : STRING := 'AlarmMgr';
	COMPONENTID : UDINT := 16#1012;
END_VAR

(* ---- DATABASEIDENTIFIERS.gvl ---- *)
VAR_GLOBAL
	TBL_ROOT_PAGES : CAA.IDENT := 8;
	IDX_ROOT_PAGES : CAA.IDENT := 2;
	IDX_ROOT_PAGES_UPDATED_FILE : CAA.IDENT := 9;
	COL_TYPE : CAA.IDENT := 0;
	COL_NAME : CAA.IDENT := 1;
	COL_TBL_NAME : CAA.IDENT := 2;
	COL_ROOTPAGE : CAA.IDENT := 3;
	COL_TIMESTAMP_LAST : CAA.IDENT := 0;
	COL_TIMESTAMP_ACTIVE : CAA.IDENT := 1;
	COL_TIMESTAMP_INACTIVE : CAA.IDENT := 2;
	COL_TIMESTAMP_ACKNOWLEDGE : CAA.IDENT := 3;
	COL_TRIGGER_VALUE : CAA.IDENT := 4;
	COL_TRIGGER_VALUE_TYPE : CAA.IDENT := 5;
	COL_LATCHVAR1_VALUE : CAA.IDENT := 6;
	COL_LATCHVAR1_TYPE : CAA.IDENT := 7;
	COL_LATCHVAR2_VALUE : CAA.IDENT := 8;
	COL_LATCHVAR2_TYPE : CAA.IDENT := 9;
	COL_GROUP_ID : CAA.IDENT := 10;
	COL_ALARM_ID : CAA.IDENT := 11;
	COL_CLASS_ID : CAA.IDENT := 12;
	COL_PRIORITY : CAA.IDENT := 13;
	COL_STATE : CAA.IDENT := 14;
	COL_OFFSET_LAST : CAA.IDENT := 15;
	COL_OFFSET_ACTIVE : CAA.IDENT := 16;
	COL_OFFSET_INACTIVE : CAA.IDENT := 17;
	COL_OFFSET_ACKNOWLEDGE : CAA.IDENT := 18;
	COL_REMOTE_DEVICE : CAA.IDENT := 19;
	COL_REMOTE_ROWID : CAA.IDENT := 20;
	COL_COMMENT_ACTIVE : CAA.IDENT := 21;
	COL_COMMENT_ACTIVEACK : CAA.IDENT := 22;
	COL_COMMENT_WAITINGCONF : CAA.IDENT := 23;
	COL_COMMENT_NORMAL : CAA.IDENT := 24;
	COL_USERID_CMT_ACTIVE : CAA.IDENT := 25;
	COL_USERID_CMT_ACTIVEACK : CAA.IDENT := 26;
	COL_USERID_CMT_WAITINGCONF : CAA.IDENT := 27;
	COL_USERID_CMT_NORMAL : CAA.IDENT := 28;
	COL_MAX_VERSION_3 : INT := ANY_TO_INT(COL_STATE);
	COL_MAX_VERSION_4 : INT := ANY_TO_INT(COL_OFFSET_ACKNOWLEDGE);
	COL_MAX_VERSION_5 : INT := ANY_TO_INT(COL_OFFSET_ACKNOWLEDGE);
	COL_MAX_VERSION_6 : INT := ANY_TO_INT(COL_REMOTE_ROWID);
	COL_MAX_VERSION_7 : INT := ANY_TO_INT(COL_USERID_CMT_NORMAL);
	COL_MAX_VERSION_DEFAULT : INT := ANY_TO_INT(COL_MAX_VERSION_7);
	COL_BYTE_ORDER : CAA.IDENT := 0;
	COL_VERSION : CAA.IDENT := 0;
	COL_LATCHVAR_VALUE : CAA.IDENT := 0;
	COL_LATCHVAR_TYPE : CAA.IDENT := 1;
END_VAR

(* ---- DBVERSIONS.gvl ---- *)
VAR_GLOBAL
	VERSION_1 : INT := 1;
	VERSION_2 : INT := 2;
	VERSION_3 : INT := 3;
	VERSION_4 : INT := 4;
	VERSION_5 : INT := 5;
	VERSION_6 : INT := 6;
	VERSION_7 : INT := 7;
	LATEST_VERSION : INT := VERSION_7;
END_VAR

(* ---- ERRORHANDLINGCONSTANTS.gvl ---- *)
VAR_GLOBAL
	METHOD_WRITE_TO_STORAGE : INT := 100;
	FUNCTION_GET_COUNT_ALARMS_FROM_STORAGE : INT := 101;
	FUNCTION_GET_ALARMS_FROM_STORAGE : INT := 102;
	METHOD_IS_RELEVANT_ALARM : INT := 103;
	FUNCTION_SKIP_ROWS : INT := 104;
	FUNCTION_GET_TIMESTAMP_VALUE : INT := 105;
	FUNCTION_POSITION_CURSOR : INT := 106;
	METHOD_CHECK_FILE_LIMIT_REACHED : INT := 107;
	METHOD_WRITE_BYTE_ORDER_FLAG : INT := 108;
	METHOD_BEGIN_TRANSACTION : INT := 109;
	METHOD_END_TRANSACTION : INT := 110;
	METHOD_SET_STATE : INT := 111;
	METHOD_DETERMINE_ROOT_PAGES : INT := 112;
	METHOD_DETERMINE_DATABASE_VERSION : INT := 113;
	METHOD_PRV_RETRIEVE_LATCH_VAR_VALUE : INT := 114;
	METHOD_CYCLIC_CALL : INT := 115;
	METHOD_ALLOCATE_ALARMGROUP_FILTER_BUFFER : INT := 116;
	METHOD_ALLOCATE_ALARMCLASS_FILTER_BUFFER : INT := 117;
	METHOD_ALLOCATE_LACTH_VARIABLES_BUFFER : INT := 118;
	METHOD_GET_MIN_MAX_TIMESTAMPS : INT := 119;
	METHOD_PRV_FIND_ROWID : INT := 120;
	METHOD_READ : INT := 121;
	METHOD_PRV_TBL_ALARM_FIND_TIMESTAMP : INT := 122;
	METHOD_BEFORE_READING : INT := 123;
	METHOD_ALLOCATE_ALARMS_TO_ACK_BUFFER : INT := 125;
	METHOD_PRV_WRITE_TO_TBL_LATCH_VAR_STRING : INT := 126;
	METHOD_PRV_OPEN_LATCH_VAR_STRINGS_TABLE_AND_CURSOR : INT := 127;
	METHOD_PRV_CLOSE_LATCH_VAR_STRINGS_TABLE_AND_CURSOR : INT := 128;
	METHOD_PRV_READ_LATCH_VAR_STRING : INT := 129;
	METHOD_PRV_ENLARGE_BUFFER_IF_NECESSARY : INT := 130;
	METHOD_PRV_SEARCH_MIN_ROW_ID : INT := 131;
	METHOD_ALLOCATE_ALARM_STORAGE_ROW_ARRAY : INT := 132;
	METHOD_CREATE_ALARM_STORAGE_METADATA_FILE : INT := 133;
	METHOD_PRV_OPEN_VERSION_TABLE : INT := 134;
	METHOD_GET_BYTE_ORDER_FLAG : INT := 135;
	METHOD_GET_FIR_LAS_ROWID : INT := 136;
	FUNCTION_GET_ALARMS_FROM_STORAGE3 : INT := 137;
	FUNCTION_GET_ALARMS_FROM_STORAGE4 : INT := 138;
	METHOD_SCAN_STORAGE : INT := 139;
	METHOD_PRV_FIND_LATCH_VAR_STRING_DBRECENT : INT := 140;
	METHOD_PRV_FIND_LATCH_VAR_STRING_DBVBEFORE5 : INT := 141;
	METHOD_PRV_FIND_LATCH_VAR_STRING : INT := 142;
	METHOD_DB_FILEWRITECONTEXT_INITIALIZE : INT := 143;
	METHOD_GETSTRINGLATCHTABLE : INT := 144;
	METHOD_DETERMINE_ROOT_PAGES_OPENSTORAGE : INT := 145;
	METHOD_GETCOUNTALLALARMSFROMSTORAGE : INT := 146;
	METHOD_DELETE_ALARMS : INT := 147;
	METHOD_CHECK_FILE_LIMIT_REACHED2 : INT := 148;
	METHOD_STORAGE_REORG : INT := 149;
	METHOD_METRICS : INT := 150;
	METHOD_SET_EMPTY_TIMESTAMP_INACTIVE : INT := 151;
	METHOD_PRV_STORE_ALARM_COMMENTS : INT := 152;
	ERRCODE_UNABLE_TO_GET_CURRENT_ROW : INT := 5;
	ACTION_SET_COL_TIMESTAMP_LAST : INT := 1000;
	ACTION_SET_COL_TIMESTAMP_ACTIVE : INT := 1001;
	ACTION_SET_COL_TIMESTAMP_INACTIVE : INT := 1002;
	ACTION_SET_COL_TIMESTAMP_ACKNOWLEDGE : INT := 1003;
	ACTION_SET_COL_TRIGGER_VALUE : INT := 1004;
	ACTION_SET_COL_LATCHVAR_VALUE : INT := 1008;
	ACTION_SET_COL_GROUP_ID : INT := 1010;
	ACTION_SET_COL_ALARM_ID : INT := 1011;
	ACTION_SET_COL_CLASS_ID : INT := 1012;
	ACTION_SET_COL_PRIORITY : INT := 1013;
	ACTION_SET_COL_STATE : INT := 1014;
	ACTION_CREATE_ROW : INT := 1015;
	ACTION_INSERT_ROW : INT := 1016;
	ACTION_SELECT_ROW : INT := 1017;
	ACTION_UPDATE_ROW : INT := 1018;
	ACTION_RELEASE_ROW : INT := 1019;
	ACTION_DELETE_ROW : INT := 1020;
	ACTION_CURSOR_OPEN : INT := 1021;
	ACTION_CURSOR_CLOSE : INT := 1022;
	ACTION_CURSOR_MOVE_FIRST : INT := 1023;
	ACTION_CURSOR_MOVE_LAST : INT := 1024;
	ACTION_CURSOR_MOVE_NEXT : INT := 1025;
	ACTION_CURSOR_MOVE_PREVIOUS : INT := 1026;
	ACTION_CURSOR_SEARCH_ROW_ID : INT := 1027;
	ACTION_CURSOR_SEARCH_INT32 : INT := 1028;
	ACTION_STORAGE_REORG : INT := 1029;
	ACTION_OPEN_TABLE : INT := 1030;
	ACTION_GET_COL_TIMESTAMP : INT := 1050;
	ACTION_GET_COL_TRIGGER_VALUE : INT := 1054;
	ACTION_GET_COL_TRIGGER_VALUE_TYPE : INT := 1055;
	ACTION_GET_COL_LATCHVAR1_VALUE : INT := 1056;
	ACTION_GET_COL_LATCHVAR1_TYPE : INT := 1057;
	ACTION_GET_COL_LATCHVAR2_VALUE : INT := 1058;
	ACTION_GET_COL_LATCHVAR2_TYPE : INT := 1059;
	ACTION_GET_COL_GROUP_ID : INT := 1060;
	ACTION_GET_COL_ALARM_ID : INT := 1061;
	ACTION_GET_COL_CLASS_ID : INT := 1062;
	ACTION_GET_COL_PRIORITY : INT := 1063;
	ACTION_GET_COL_STATE : INT := 1064;
	ACTION_SET_COL_BYTE_ORDER : INT := 1065;
	ACTION_STORAGE_OPEN : INT := 1066;
	ACTION_BEGIN_TRANSACTION : INT := 1067;
	ACTION_END_TRANSACTION : INT := 1068;
	ACTION_GET_COL_VERSION : INT := 1069;
	ACTION_TEXT_COPY_TO_STRING : INT := 1070;
	ACTION_GET_COL_TYPE : INT := 1071;
	ACTION_GET_COL_NAME : INT := 1072;
	ACTION_GET_COL_TBL_NAME : INT := 1073;
	ACTION_GET_COL_ROOTPAGE : INT := 1074;
	ACTION_GET_COL_LATCHVAR_VALUE : INT := 1075;
	ACTION_GET_COL_LATCHVAR_TYPE : INT := 1076;
	ACTION_CURSOR_CURRENT_ROW : INT := 1077;
	ACTION_TABLE_NUM_OF_ROWS : INT := 1078;
	ACTION_TABLE_GET_MINMAXROWIDS : INT := 1079;
	ACTION_GET_COL_OFFSET_LAST : INT := 1080;
	ACTION_GET_COL_OFFSET_ACTIVE : INT := 1081;
	ACTION_GET_COL_OFFSET_INACTIVE : INT := 1082;
	ACTION_GET_COL_OFFSET_ACKNOWLEDGE : INT := 1083;
	ACTION_SET_COL_OFFSET_LAST : INT := 1084;
	ACTION_SET_COL_OFFSET_ACTIVE : INT := 1085;
	ACTION_SET_COL_OFFSET_INACTIVE : INT := 1086;
	ACTION_SET_COL_OFFSET_ACKNOWLEDGE : INT := 1087;
	ACTION_GET_COL_BYTE_ORDER : INT := 1088;
	ACTION_SET_COL_DEVICE_NAME : INT := 1089;
	ACTION_SET_COL_DEVICE_ROWID : INT := 1090;
	ACTION_GET_COL_DEVICE_NAME : INT := 1091;
	ACTION_GET_COL_DEVICE_ROWID : INT := 1092;
	ACTION_GET_COL_TIMESTAMP_ACTIVE : INT := 1093;
	ACTION_CURSOR_SEARCH_TEXT : INT := 1094;
	ACTION_STORAGE_OPEN_ROLLBACKATTEMPT : INT := 1095;
	ACTION_METRICS : INT := 1096;
	ACTION_SET_COL_CMT_ACTIVE : INT := 1097;
	ACTION_SET_COL_CMT_ACTIVEACK : INT := 1098;
	ACTION_SET_COL_CMT_WAITINGCONF : INT := 1099;
	ACTION_SET_COL_CMT_NORMAL : INT := 1100;
	ACTION_SET_COL_USERID_ACTIVE : INT := 1101;
	ACTION_SET_COL_USERID_ACTIVEACK : INT := 1102;
	ACTION_SET_COL_USERID_WAITINGCONF : INT := 1103;
	ACTION_SET_COL_USERID_NORMAL : INT := 1104;
	ACTION_GET_COL_CMT_ACTIVE : INT := 1105;
	ACTION_GET_COL_CMT_ACTIVEACK : INT := 1106;
	ACTION_GET_COL_CMT_WAITINGCONF : INT := 1107;
	ACTION_GET_COL_CMT_NORMAL : INT := 1108;
	ACTION_GET_COL_USERID_ACTIVE : INT := 1109;
	ACTION_GET_COL_USERID_ACTIVEACK : INT := 1110;
	ACTION_GET_COL_USERID_WAITINGCONF : INT := 1111;
	ACTION_GET_COL_USERID_NORMAL : INT := 1112;
	ACTION_CREATE_TEXT_FROM_STRING : INT := 3060;
	ACTION_TEXT_FREE : INT := 3061;
END_VAR

(* ---- EVENTS.gvl ---- *)
VAR_GLOBAL
	EVT_ALARMMANAGERGETCOUNT : UDINT := 16#10001;
	EVT_ALARMMANAGERGETALARMS : UDINT := 16#10002;
	EVT_ALARMMANAGERHANDLESERVICE : UDINT := 16#10003;
	EVT_CHSCHANNELCLOSED : UDINT := 16#10001;
	CMPID_CMPCHANNELSERVER : UDINT := 16#A;
	CMPID_CMPALARMMANAGER : UDINT := 16#7C;
	INVALID_HANDLE : RTS_IEC_HANDLE := 16#FFFFFFFF;
	RETVAL_OK : UINT := 16#0;
	RETVAL_BUFFEROVERFLOW : UINT := 16#2;
	EVT_LOC_CHANNEL_CLOSED : INT := 1;
END_VAR

(* ---- GLOBALLYFORALARMSTORAGE.gvl ---- *)
VAR_GLOBAL
	G_EVENTDISPATCHER : EventDispatcher;
	G_ALARMSTORAGEMANAGER : AlarmStorageManager;
	G_ALARMSTORAGEREADER : AlarmStorageReader;
	G_SQLITEDATABASEACCESS : SQLiteDatabaseAccess;
	G_ALARMSTORAGEREADERCONSUMER : AlarmServiceAlarmStorageReaderConsumer;
	G_ROOTPAGEREADWRITEMODEPROVIDER : AlarmRootPageReadWriteModeProvider;
	G_BDUMMY : BOOL;
END_VAR

(* ---- MONITOR.gvl ---- *)
VAR_GLOBAL
	FILTERBYLATCH : MonitorFilterByLatch;
	FILTERBYDATETIME : MonitorFilterByDateTime;
	DBSTATUS : MonitorDBStatus;
	COMPILECHECKONLY : BOOL;
END_VAR

(* ---- PROXYCONSTANTS.gvl ---- *)
VAR_GLOBAL
	REQ_ID_NONE : INT := -1;
	REQ_ID_GET_DEVICE_NAME : INT := 1;
	REQ_ID_GET_LATCHVARS_COUNT : INT := 2;
	REQ_ID_GET_TOTALM_COUNT : INT := 3;
	REQ_ID_GET_TOTCLA_COUNT : INT := 4;
	REQ_ID_SET_HIST_ALARM_RECORD : INT := 5;
	REQ_ID_SET_ALARM_RECORD : INT := 10;
	REQ_ID_RES_ALARM_RECORD : INT := 11;
	REQ_ID_READ_ACTIVE_ALARMS : INT := 12;
	REQ_ID_READ_ALARMS_CONFIG : INT := 13;
	REQ_ID_READ_CLASS_CONFIG : INT := 14;
	REQ_ID_ACK_ALARMS : INT := 15;
	REQ_ID_READ_HIST_CONFIG : INT := 16;
	REQ_ID_READ_HIST_ALARMS : INT := 17;
	REQ_ID_READ_HIST_ACTIVE_ALARMS : INT := 18;
	REQ_ID_CHANNEL_TEST : INT := 100;
	REQ_ID_CHANNEL_TEST2 : INT := 101;
	FIFO_ERROR_SIZE : INT := 10;
	AREQID : ARRAY [1..MAX_TASK_TEST] OF INT := [REQ_ID_CHANNEL_TEST, REQ_ID_CHANNEL_TEST2, REQ_ID_SET_ALARM_RECORD, REQ_ID_RES_ALARM_RECORD, REQ_ID_READ_ACTIVE_ALARMS, REQ_ID_READ_ALARMS_CONFIG, REQ_ID_READ_CLASS_CONFIG, REQ_ID_ACK_ALARMS, REQ_ID_READ_HIST_CONFIG, REQ_ID_READ_HIST_ALARMS, REQ_ID_READ_HIST_ACTIVE_ALARMS];
	MAX_TASK : INT := 7;
	MAX_TASK_TEST : INT := 11;
END_VAR

(* ---- PROXYGVL.gvl ---- *)
VAR_GLOBAL
	PROXYALLOC : Allocator;
END_VAR

(* ---- RETURNVALUES.gvl ---- *)
VAR_GLOBAL
	ERR_OK : UDINT := Errors.ERR_OK;
	ERR_NOTINITIALIZED : UDINT := Errors.ERR_NOTINITIALIZED;
	ERR_PARAMETER : UDINT := Errors.ERR_PARAMETER;
	ERR_NO_OBJECT : UDINT := Errors.ERR_NO_OBJECT;
	ERR_DUPLICATE : UDINT := Errors.ERR_DUPLICATE;
	ERR_NO_ALARM_MANAGER_CLIENT : UDINT := 16#1000;
	ERR_NO_FILTER_CRITERIA : UDINT := 16#1001;
	ERR_NO_ALARMGROUP_FILTER_CRITERIA : UDINT := 16#1002;
	ERR_NO_ALARMCLASS_FILTER_CRITERIA : UDINT := 16#1003;
	ERR_INVALID_PRIORITY_FILTER : UDINT := 16#1004;
	ERR_NO_ALARM_STORAGE : UDINT := 16#1005;
	ERR_UNEXPECTED_ALARMSTATE : UDINT := 16#1006;
END_VAR

(* ---- IACKALARMSSERVICECONSUMER.itf ---- *)
INTERFACE IACKALARMSSERVICECONSUMER
END_INTERFACE

(* ---- IACKALARMSSERVICEPROVIDER.itf ---- *)
INTERFACE IACKALARMSSERVICEPROVIDER
END_INTERFACE

METHOD GETCOUNTALARMSTOACKNOWLEDGE : INT
END_METHOD

METHOD GETNEXTALARMTOACKNOWLEDGE : BOOL
VAR_INPUT
	XFISRTENTRY : BOOL;
END_VAR
VAR_OUTPUT
	ALARMTOACKNOWLEDGE : AlarmToAcknowledge;
END_VAR
END_METHOD

(* ---- IALARM.itf ---- *)
INTERFACE IALARM
END_INTERFACE

METHOD GETALARMCLASS : IAlarmClass
END_METHOD

METHOD GETALARMGROUP : IAlarmGroup
END_METHOD

METHOD GETID : ALARM_ID
END_METHOD

METHOD GETINTERNALID : UDINT
END_METHOD

METHOD GETMESSAGE : CharBufferPtr
VAR_INPUT
	STRINGTYPE : __SYSTEM.TYPE_CLASS;
END_VAR
END_METHOD

METHOD GETOBSERVATIONTYPE : IAlarmObservationType
END_METHOD

METHOD GETROWID : CAA.IDENT
END_METHOD

METHOD GETSTATE : AlarmState
END_METHOD

METHOD ISDEACTIVATED : BOOL
END_METHOD

METHOD SETALARMCLASS
VAR_INPUT
	ITFALARMCLASS : IAlarmClass;
END_VAR
END_METHOD

METHOD SETALARMGROUP
VAR_INPUT
	ITFALARMGROUP : IAlarmGroup;
END_VAR
END_METHOD

METHOD SETHIGHERPRIOALARM
VAR_INPUT
	ITFALARM : IAlarm;
END_VAR
END_METHOD

METHOD SETOBSERVATIONTYPE
VAR_INPUT
	ITFOBSERVATIONTYPE : IAlarmObservationType;
END_VAR
END_METHOD

METHOD SETROWID
VAR_INPUT
	ROWID : CAA.IDENT;
END_VAR
END_METHOD

METHOD SETTIMESTAMP
VAR_INPUT
	LICURRTIMESTAMP : Timestamp;
	ESTATE : AlarmState;
	ESTATETRANSITION : AlarmStateTransition;
END_VAR
END_METHOD

METHOD GETTIMESTAMPACKNOWLEDGE : Timestamp
END_METHOD

METHOD GETTIMESTAMPACTIVE : Timestamp
END_METHOD

METHOD GETTIMESTAMPINACTIVE : Timestamp
END_METHOD

METHOD GETTIMESTAMPLAST : Timestamp
END_METHOD

METHOD GETCURRENTVALUE : ITypedValue
END_METHOD

METHOD GETLATCHVAR1VALUE : ITypedValue
END_METHOD

METHOD GETLATCHVAR2VALUE : ITypedValue
END_METHOD

METHOD GETTRIGGERVALUE : ITypedValue
END_METHOD

(* ---- IALARM2.itf ---- *)
INTERFACE IALARM2
END_INTERFACE

METHOD SETALARMSTATE
VAR_INPUT
	EALARMSTATE : AlarmState;
END_VAR
END_METHOD

METHOD SETCURRENTVALUE
VAR_INPUT
	ITFTYPEDVALUECURRENT : ITypedValue;
END_VAR
END_METHOD

METHOD SETID
VAR_INPUT
	UIID : ALARM_ID;
END_VAR
END_METHOD

METHOD SETINTERNALID
VAR_INPUT
	UDIID : UDINT;
END_VAR
END_METHOD

METHOD SETLATCHVAR1VALUE
VAR_INPUT
	ITFTYPEDVALUELATCHVAR1 : ITypedValue;
END_VAR
END_METHOD

METHOD SETLATCHVAR2VALUE
VAR_INPUT
	ITFTYPEDVALUELATCHVAR2 : ITypedValue;
END_VAR
END_METHOD

METHOD SETTIMESTAMPACKNOWLEDGE
VAR_INPUT
	LITIMESTAMPACKNOWLEDGE : Timestamp;
END_VAR
END_METHOD

METHOD SETTIMESTAMPACTIVE
VAR_INPUT
	LITIMESTAMPACTIVE : Timestamp;
END_VAR
END_METHOD

METHOD SETTIMESTAMPINACTIVE
VAR_INPUT
	LITIMESTAMPINACTIVE : Timestamp;
END_VAR
END_METHOD

METHOD SETTIMESTAMPLAST
VAR_INPUT
	LITIMESTAMPLAST : Timestamp;
END_VAR
END_METHOD

METHOD SETTRIGGERVALUE
VAR_INPUT
	ITFTYPEDVALUETRIGGER : ITypedValue;
END_VAR
END_METHOD

(* ---- IALARM3.itf ---- *)
INTERFACE IALARM3
END_INTERFACE

METHOD GETCOUNTLATCHVARIABLES : USINT
END_METHOD

METHOD GETCOUNTMESSAGES : USINT
END_METHOD

METHOD GETLATCHVARVALUE : ITypedValue
VAR_INPUT
	IWHICHLATCHVAR : INT;
END_VAR
END_METHOD

METHOD GETMESSAGE2 : CharBufferPtr
VAR_INPUT
	STRINGTYPE : __SYSTEM.TYPE_CLASS;
	IWHICHMESSAGE : INT;
END_VAR
END_METHOD

METHOD SETLATCHVARVALUE
VAR_INPUT
	IWHICHLATCHVAR : INT;
	ITFTYPEDVALUELATCHVAR : ITypedValue;
END_VAR
END_METHOD

(* ---- IALARM4.itf ---- *)
INTERFACE IALARM4
END_INTERFACE

(* ---- IALARM5.itf ---- *)
INTERFACE IALARM5
END_INTERFACE

METHOD SETTIMESTAMP2
VAR_INPUT
	LICURRTIMESTAMP : Timestamp;
	IOFFSET : INT;
	ESTATE : AlarmState;
	ESTATETRANSITION : AlarmStateTransition;
END_VAR
END_METHOD

(* ---- IALARM6.itf ---- *)
INTERFACE IALARM6
END_INTERFACE

(* ---- IALARM7.itf ---- *)
INTERFACE IALARM7
END_INTERFACE

(* ---- IALARM8.itf ---- *)
INTERFACE IALARM8
END_INTERFACE

METHOD SETACKNOWLEDGE : BOOL
VAR_INPUT
	PWSCOMMENT : POINTER TO WSTRING;
	PWSUSERID : POINTER TO WSTRING;
END_VAR
END_METHOD

(* ---- IALARMADAPTER.itf ---- *)
INTERFACE IALARMADAPTER
END_INTERFACE

METHOD INITIALIZE
END_METHOD

(* ---- IALARMAPIOBSERVATIONTYPE.itf ---- *)
INTERFACE IALARMAPIOBSERVATIONTYPE
END_INTERFACE

(* ---- IALARMCLASS.itf ---- *)
INTERFACE IALARMCLASS
END_INTERFACE

METHOD GETACKNOWLEDGEMETHOD : AcknowledgeMethod
END_METHOD

METHOD GETALARMSTATEMACHINE : IAlarmStateMachine
END_METHOD

METHOD GETDISPLAYOPTIONS : POINTER TO DisplayOptions
VAR_INPUT
	ESTATE : AlarmState;
END_VAR
END_METHOD

METHOD GETINTERNALID : UDINT
END_METHOD

METHOD GETNAME : STRING
END_METHOD

METHOD GETPRIORITY : USINT
END_METHOD

METHOD ISACKNOWLEDGESEPARATELY : BOOL
END_METHOD

(* ---- IALARMCLASS2.itf ---- *)
INTERFACE IALARMCLASS2
END_INTERFACE

METHOD ACKINSTEADOFCONFIRM : BOOL
END_METHOD

METHOD AUTORESETDIGITALALARMS : BOOL
END_METHOD

(* ---- IALARMCLASS3.itf ---- *)
INTERFACE IALARMCLASS3
END_INTERFACE

METHOD GETALARMCLASSOBJECTCHECKSUM : LINT
END_METHOD

(* ---- IALARMCLASSINTERNAL.itf ---- *)
INTERFACE IALARMCLASSINTERNAL
END_INTERFACE

METHOD GETARCHIVING : BOOL
END_METHOD

METHOD NOTIFYNOTIFIABLES
VAR_INPUT
	ESTATETRANSITION : AlarmStateTransition;
	ITFALARM : IAlarm;
END_VAR
END_METHOD

(* ---- IALARMCONFIGURATION.itf ---- *)
INTERFACE IALARMCONFIGURATION
END_INTERFACE

METHOD ACKNOWLEDGEALL
END_METHOD

METHOD ACKNOWLEDGEALLOFGROUP
VAR_INPUT
	USIALARMGROUPID : ALARMGROUP_ID;
END_VAR
END_METHOD

METHOD ACKNOWLEDGEONEOFGROUP
VAR_INPUT
	USIALARMGROUPID : ALARMGROUP_ID;
	UIALARMID : ALARM_ID;
END_VAR
END_METHOD

METHOD CYCLICCALL
END_METHOD

METHOD FINDALARM : POINTER TO Alarm
VAR_INPUT
	SALARMGROUP : STRING;
	UIALARMID : ALARM_ID;
END_VAR
END_METHOD

METHOD FINDALARMCLASS : IAlarmClass
VAR_INPUT
	UDIID : UDINT;
END_VAR
END_METHOD

METHOD FINDALARMGROUP : IAlarmGroup
VAR_INPUT
	UDIID : UDINT;
END_VAR
END_METHOD

METHOD GETSTORAGE : IDatabaseFileAlarmStorage
END_METHOD

METHOD HASSTORAGE : BOOL
END_METHOD

METHOD RAISEEVENT : BOOL
VAR_INPUT
	EVENT : AlarmEvent;
END_VAR
END_METHOD

(* ---- IALARMCONFIGURATION2.itf ---- *)
INTERFACE IALARMCONFIGURATION2
END_INTERFACE

METHOD DETERMINERELEVANTALARMS : UDINT
VAR_INPUT
	ITFALARMFILTERCRITERIA : IAlarmFilterCriteria;
	PARRITFRELEVANTALARMS : POINTER TO ARRAY [0..0] OF IAlarm;
	IOFFSET : INT;
END_VAR
END_METHOD

METHOD FINDALARMGROUPBYNAME : IAlarmGroup
VAR_INPUT
	SALARMGROUP : STRING;
END_VAR
END_METHOD

(* ---- IALARMCONFIGURATION3.itf ---- *)
INTERFACE IALARMCONFIGURATION3
END_INTERFACE

METHOD FINDALARMCLASSBYNAME : IAlarmClass
VAR_INPUT
	SALARMCLASS : STRING;
END_VAR
END_METHOD

(* ---- IALARMCONFIGURATION4.itf ---- *)
INTERFACE IALARMCONFIGURATION4
END_INTERFACE

METHOD RAISEEVENT2 : BOOL
VAR_INPUT
	EVENT : AlarmEvent;
END_VAR
VAR_OUTPUT
	ITFALARM : IAlarm;
END_VAR
END_METHOD

(* ---- IALARMCONFIGURATION5.itf ---- *)
INTERFACE IALARMCONFIGURATION5
END_INTERFACE

METHOD GETALARMGROUPS : POINTER TO ARRAY [0..0] OF IAlarmGroup
VAR_OUTPUT
	IALARMGROUPCOUNT : INT;
END_VAR
END_METHOD

(* ---- IALARMCONFIGURATION6.itf ---- *)
INTERFACE IALARMCONFIGURATION6
END_INTERFACE

METHOD FINDALARMCLASSCOUNT : INT
END_METHOD

(* ---- IALARMCONFIGURATION7.itf ---- *)
INTERFACE IALARMCONFIGURATION7
END_INTERFACE

METHOD CLEARHISTORY : BOOL
VAR_INPUT
	XKEEPACTIVEALARMS : BOOL;
END_VAR
END_METHOD

(* ---- IALARMCONFIGURATION8.itf ---- *)
INTERFACE IALARMCONFIGURATION8
END_INTERFACE

(* ---- IALARMCONFIGURATION9.itf ---- *)
INTERFACE IALARMCONFIGURATION9
END_INTERFACE

METHOD ACKNOWLEDGEALLOFGROUPWITHCOMMENT
VAR_INPUT
	USIALARMGROUPID : ALARMGROUP_ID;
END_VAR
VAR_IN_OUT
	WSCOMMENT : WSTRING;
	WSUSERID : WSTRING;
END_VAR
END_METHOD

METHOD ACKNOWLEDGEALLWITHCOMMENT
VAR_IN_OUT
	WSCOMMENT : WSTRING;
	WSUSERID : WSTRING;
END_VAR
END_METHOD

METHOD ACKNOWLEDGEONEOFGROUPWITHCOMMENT
VAR_INPUT
	USIALARMGROUPID : ALARMGROUP_ID;
	UIALARMID : ALARM_ID;
END_VAR
VAR_IN_OUT
	WSCOMMENT : WSTRING;
	WSUSERID : WSTRING;
END_VAR
END_METHOD

METHOD SETCOMMENT : UDINT
VAR_INPUT
	USIALARMGROUPID : ALARMGROUP_ID;
	UIALARMID : ALARM_ID;
END_VAR
VAR_IN_OUT
	WSCOMMENT : WSTRING;
	WSUSERID : WSTRING;
END_VAR
END_METHOD

(* ---- IALARMCONFIGURATIONREMOTE.itf ---- *)
INTERFACE IALARMCONFIGURATIONREMOTE
END_INTERFACE

METHOD CYCLICCALL
END_METHOD

METHOD GETACTIVEALARMS
VAR_INPUT
	PASNAME : POINTER TO ARRAY [0..10] OF STRING;
	IGROUPCOUNT : INT;
	FILTERCRITERIA : REFERENCE TO VisuFbAlarmFilterCriteria;
	ITFALARMDATABLOCK : IAlarmDataBlockBaseDINT;
END_VAR
VAR_IN_OUT
	DISTUBPROG : DINT;
END_VAR
END_METHOD

METHOD GETALARMCLASSDESC : BOOL
VAR_INPUT
	SPROXYNAME : STRING;
	UDIID : UDINT;
END_VAR
VAR_OUTPUT
	SDESC : ProxyStructAlarmClassDesc;
END_VAR
END_METHOD

METHOD GETALARMCLASSDESCBYNAME : BOOL
VAR_INPUT
	SPROXYNAME : STRING;
	SCLASSNAME : STRING;
END_VAR
VAR_OUTPUT
	SDESC : ProxyStructAlarmClassDesc;
END_VAR
END_METHOD

METHOD GETALARMDESC : BOOL
VAR_INPUT
	SPROXYNAME : STRING;
	UDIALMID : UDINT;
	UDIGRPID : UDINT;
END_VAR
VAR_OUTPUT
	SDESC : ProxyStructAlarmDesc;
END_VAR
END_METHOD

METHOD GETALARMDISPLAYOPTIONS : BOOL
VAR_INPUT
	ITFALARMMETAOBJECTSTUB5 : IAlarmMetaObjectStub5;
	REFDISPLAYOPTIONS : REFERENCE TO DisplayOptions;
END_VAR
VAR_OUTPUT
	XVALID : BOOL;
	SCLASSREMAP : STRING;
END_VAR
END_METHOD

METHOD GETALARMGROUPDESC : BOOL
VAR_INPUT
	SPROXYNAME : STRING;
	UDIID : UDINT;
END_VAR
VAR_OUTPUT
	SDESC : ProxyStructAlarmGroupDesc;
END_VAR
END_METHOD

METHOD GETALARMGROUPDESCBYNAME : BOOL
VAR_INPUT
	SPROXYNAME : STRING;
	SGRPNAME : STRING;
END_VAR
VAR_OUTPUT
	SDESC : ProxyStructAlarmGroupDesc;
END_VAR
END_METHOD

METHOD GETALARMMESSAGE : BOOL
VAR_INPUT
	ITFALARMMETAOBJECTSTUB5 : IAlarmMetaObjectStub5;
	IWHICHMESSAGE : INT;
	REFCHARBUFFERSTRING : REFERENCE TO CharBufferString;
	STRINGTYPE : __SYSTEM.TYPE_CLASS;
END_VAR
END_METHOD

METHOD GETALARMMESSAGE2 : BOOL
VAR_INPUT
	SNAME : STRING;
	STEXTLISTNAME : STRING;
	STEXTLISTINDEX : STRING;
	IWHICHMESSAGE : INT;
	STRINGTYPE : __SYSTEM.TYPE_CLASS;
END_VAR
VAR_OUTPUT
	MESSAGE : CharBufferPtr;
END_VAR
END_METHOD

METHOD GETPROXY : IProxy
VAR_INPUT
	SNAME : STRING;
END_VAR
END_METHOD

METHOD GETPROXYALARMCLASSESDESCRIPTION : BOOL
VAR_INPUT
	SNAME : STRING;
	PCLDESC : POINTER TO ARRAY [0..0] OF ProxyStructMonitorAlarmClassDesc;
	ISIZE : INT;
END_VAR
VAR_OUTPUT
	ICLCNT : INT;
END_VAR
END_METHOD

METHOD GETPROXYALARMGROUPSDESCRIPTION : BOOL
VAR_INPUT
	SNAME : STRING;
	PGRPDESC : POINTER TO ARRAY [0..0] OF ProxyStructMonitorAlarmGroupDesc;
	ISIZE : INT;
END_VAR
VAR_OUTPUT
	IGRPCNT : INT;
END_VAR
END_METHOD

METHOD GETPROXYALARMSDESCRIPTION : BOOL
VAR_INPUT
	SNAME : STRING;
	PALMDESC : POINTER TO ARRAY [0..0] OF ProxyStructMonitorAlarmDesc;
	DISIZE : DINT;
END_VAR
VAR_OUTPUT
	DIALMCNT : DINT;
END_VAR
END_METHOD

METHOD GETPROXYSTATISTICS : BOOL
VAR_INPUT
	SNAME : STRING;
END_VAR
VAR_OUTPUT
	STRUCTMONITOR : ProxyStructMonitor;
END_VAR
END_METHOD

METHOD GETPROXYSTATISTICSSINGLEACTIVITY : BOOL
VAR_INPUT
	SNAME : STRING;
	ITASKID : INT;
END_VAR
VAR_OUTPUT
	STRUCTMONITOR : ProxyStructMonitorRequest;
END_VAR
END_METHOD

METHOD GETSTORAGE : IDatabaseFileAlarmStorage
END_METHOD

METHOD HASSTORAGE : BOOL
END_METHOD

METHOD REGISTERUSERCLIENT : BOOL
VAR_INPUT
	IINDEX : INT;
END_VAR
VAR_OUTPUT
	ITFPROXY : IProxy;
END_VAR
END_METHOD

METHOD SETALARMSTOACK
VAR_INPUT
	ITFALARMDATABLOCK : IAlarmDataBlockBase2;
END_VAR
END_METHOD

(* ---- IALARMCONFIGURATIONSUPPORTSTRAVERSAL.itf ---- *)
INTERFACE IALARMCONFIGURATIONSUPPORTSTRAVERSAL
END_INTERFACE

METHOD TRAVERSEALLALARMSOFALLALARMGROUPS
VAR_INPUT
	ITFALARMTRAVERSALCONSUMER : IAlarmTraversalConsumer;
END_VAR
END_METHOD

METHOD TRAVERSEALLCLASSES
VAR_INPUT
	ITFALARMTRAVERSALCONSUMER : IAlarmTraversalConsumer;
END_VAR
END_METHOD

(* ---- IALARMGROUP.itf ---- *)
INTERFACE IALARMGROUP
END_INTERFACE

METHOD FINDALARM : POINTER TO Alarm
VAR_INPUT
	UDIID : UDINT;
END_VAR
END_METHOD

METHOD FINDALARM2 : POINTER TO Alarm
VAR_INPUT
	UIID : ALARM_ID;
END_VAR
END_METHOD

METHOD GETALARMSTORAGE : IDatabaseFileAlarmStorage
END_METHOD

METHOD GETALARMS : POINTER TO ARRAY [0..0] OF Alarm
VAR_OUTPUT
	IALARMCOUNT : INT;
END_VAR
END_METHOD

METHOD GETEVENTS : POINTER TO ARRAY [0..0] OF Alarm
VAR_OUTPUT
	IEVENTCOUNT : INT;
END_VAR
END_METHOD

METHOD GETINTERNALID : UDINT
END_METHOD

METHOD GETNAME : STRING
END_METHOD

METHOD GETSTRINGID : STRING
VAR_INPUT
	UIID : ALARM_ID;
END_VAR
END_METHOD

METHOD GETTEXTLISTNAME : POINTER TO STRING
END_METHOD

METHOD GETVALUEPROVIDER : IValueProvider
END_METHOD

METHOD ISDEACTIVATED : BOOL
END_METHOD

METHOD RAISEEVENT : BOOL
VAR_INPUT
	EVENT : AlarmEvent;
END_VAR
END_METHOD

METHOD SETACTIVEALARM
VAR_INPUT
	IINDEX : INT;
	PALARM : POINTER TO Alarm;
END_VAR
END_METHOD

METHOD SETACTIVEALARMCOUNT
VAR_INPUT
	ICOUNT : INT;
END_VAR
END_METHOD

(* ---- IALARMGROUP2.itf ---- *)
INTERFACE IALARMGROUP2
END_INTERFACE

METHOD GETTEXTID : STRING
VAR_INPUT
	UIID : ALARM_ID;
	IWHICHMESSAGE : INT;
END_VAR
END_METHOD

(* ---- IALARMGROUP3.itf ---- *)
INTERFACE IALARMGROUP3
END_INTERFACE

METHOD GETID : ALARMGROUP_ID
END_METHOD

METHOD SETID
VAR_INPUT
	USIALARMGROUPID : ALARMGROUP_ID;
END_VAR
END_METHOD

(* ---- IALARMGROUP4.itf ---- *)
INTERFACE IALARMGROUP4
END_INTERFACE

METHOD GETSTRINGID2 : STRING
VAR_INPUT
	UDIALARMID : UDINT;
	IWHICHMESSAGE : INT;
END_VAR
VAR_OUTPUT
	STEXTID : STRING;
END_VAR
END_METHOD

(* ---- IALARMGROUP5.itf ---- *)
INTERFACE IALARMGROUP5
END_INTERFACE

METHOD RAISEEVENT2 : BOOL
VAR_INPUT
	EVENT : AlarmEvent;
END_VAR
VAR_OUTPUT
	ITFALARM : IAlarm;
END_VAR
END_METHOD

(* ---- IALARMGROUP6.itf ---- *)
INTERFACE IALARMGROUP6
END_INTERFACE

METHOD GETTEXTLISTNAME2 : POINTER TO STRING
VAR_INPUT
	UIID : ALARM_ID;
END_VAR
END_METHOD

(* ---- IALARMGROUPSUPPORTSTRAVERSAL.itf ---- *)
INTERFACE IALARMGROUPSUPPORTSTRAVERSAL
END_INTERFACE

METHOD TRAVERSEALLALARMS
VAR_INPUT
	IWHICHALARMGROUP : INT;
	ITFALARMTRAVERSALCONSUMER : IAlarmTraversalConsumer;
END_VAR
END_METHOD

(* ---- IALARMHANDLER.itf ---- *)
INTERFACE IALARMHANDLER
END_INTERFACE

METHOD ACKNOWLEDGEALL
END_METHOD

METHOD ACKNOWLEDGEALLOFGROUP
VAR_INPUT
	USIALARMGROUPID : ALARMGROUP_ID;
END_VAR
END_METHOD

METHOD ACKNOWLEDGEONEOFGROUP
VAR_INPUT
	USIALARMGROUPID : ALARMGROUP_ID;
	UIALARMID : ALARM_ID;
END_VAR
END_METHOD

METHOD CYCLICCALL
END_METHOD

METHOD FINDALARMCLASS : IAlarmClass
VAR_INPUT
	UDIID : UDINT;
END_VAR
END_METHOD

METHOD FINDALARMGROUP : IAlarmGroup
VAR_INPUT
	UDIID : UDINT;
END_VAR
END_METHOD

METHOD GETSTORAGE : IDatabaseFileAlarmStorage
END_METHOD

METHOD HASSTORAGE : BOOL
END_METHOD

METHOD RAISEEVENT : BOOL
VAR_INPUT
	USIALARMGROUPID : ALARMGROUP_ID;
	UIALARMID : ALARM_ID;
END_VAR
END_METHOD

METHOD REGISTERALARMCONFIGURATION
VAR_INPUT
	ITFALARMCONFIGURATION : IAlarmConfiguration;
END_VAR
END_METHOD

(* ---- IALARMHANDLER2.itf ---- *)
INTERFACE IALARMHANDLER2
END_INTERFACE

METHOD GETACTIVEALARMS : UDINT
VAR_INPUT
	ITFALARMMANAGERCLIENT : IAlarmManagerClient;
END_VAR
VAR_OUTPUT
	PARRITFACTIVEALARMS : POINTER TO ARRAY [0..0] OF IAlarm;
	ICOUNTACTIVEALARMS : INT;
END_VAR
END_METHOD

METHOD GETALARMSFROMSTORAGE : UDINT
VAR_INPUT
	ITFALARMMANAGERCLIENT : IAlarmManagerClient;
	ISKIPROWS : INT;
END_VAR
VAR_OUTPUT
	ICOUNTROWS : INT;
END_VAR
VAR_IN_OUT
	BROWIDVALID : BOOL;
	DIROWID : DINT;
END_VAR
END_METHOD

METHOD GETCOUNTALARMSFROMSTORAGE : DINT
VAR_INPUT
	ITFALARMMANAGERCLIENT : IAlarmManagerClient;
END_VAR
VAR_OUTPUT
	UDIRESULT : UDINT;
END_VAR
END_METHOD

METHOD REGISTERCLIENT : UDINT
VAR_INPUT
	ITFALARMMANAGERCLIENT : IAlarmManagerClient;
	PARRITFALARMSFROMHISTORY : POINTER TO ARRAY [0..0] OF IAlarm2;
	ICOUNTALARMSFROMHISTORY : INT;
END_VAR
END_METHOD

METHOD UNREGISTERCLIENT : UDINT
VAR_INPUT
	ITFALARMMANAGERCLIENT : IAlarmManagerClient;
END_VAR
END_METHOD

(* ---- IALARMHANDLER3.itf ---- *)
INTERFACE IALARMHANDLER3
END_INTERFACE

METHOD UNREGISTERALARMCONFIGURATION
VAR_INPUT
	ITFALARMCONFIGURATION : IAlarmConfiguration;
END_VAR
END_METHOD

(* ---- IALARMHANDLER4.itf ---- *)
INTERFACE IALARMHANDLER4
END_INTERFACE

METHOD REGISTERALARMSTATECHANGEDLISTENER : BOOL
VAR_INPUT
	ITFALARMSTATECHANGEDLISTENER : IAlarmStateChangedListener;
END_VAR
END_METHOD

(* ---- IALARMHANDLER5.itf ---- *)
INTERFACE IALARMHANDLER5
END_INTERFACE

METHOD GETALARMCONFIGURATION : IAlarmConfiguration
VAR_INPUT
	IPOS : INT;
END_VAR
END_METHOD

(* ---- IALARMHANDLER6.itf ---- *)
INTERFACE IALARMHANDLER6
END_INTERFACE

METHOD ACKNOWLEDGEALLOFGROUPWITHCOMMENT
VAR_INPUT
	USIALARMGROUPID : ALARMGROUP_ID;
END_VAR
VAR_IN_OUT
	WSCOMMENT : WSTRING;
	WSUSERID : WSTRING;
END_VAR
END_METHOD

METHOD ACKNOWLEDGEALLWITHCOMMENT
VAR_IN_OUT
	WSCOMMENT : WSTRING;
	WSUSERID : WSTRING;
END_VAR
END_METHOD

METHOD ACKNOWLEDGEONEOFGROUPWITHCOMMENT
VAR_INPUT
	USIALARMGROUPID : ALARMGROUP_ID;
	UIALARMID : ALARM_ID;
END_VAR
VAR_IN_OUT
	WSCOMMENT : WSTRING;
	WSUSERID : WSTRING;
END_VAR
END_METHOD

METHOD SETCOMMENT : UDINT
VAR_INPUT
	USIALARMGROUPID : ALARMGROUP_ID;
	UIALARMID : ALARM_ID;
END_VAR
VAR_IN_OUT
	WSCOMMENT : WSTRING;
	WSUSERID : WSTRING;
END_VAR
END_METHOD

(* ---- IALARMHANDLER7.itf ---- *)
INTERFACE IALARMHANDLER7
END_INTERFACE

METHOD GETINSTANCEALARM : IAlarm8
VAR_INPUT
	PFBINSTANCE : POINTER TO BYTE;
	UITEMPLATEALARMID : ALARM_ID;
END_VAR
VAR_OUTPUT
	USIALARMGROUPID : ALARMGROUP_ID;
	UIALARMID : ALARM_ID;
END_VAR
END_METHOD

METHOD GETINSTANCEALARMBYNAME : IAlarm8
VAR_INPUT
	PFBINSTANCE : POINTER TO BYTE;
	UITEMPLATEALARMID : ALARM_ID;
	STALARMTEMPLATENAME : STRING(255);
END_VAR
VAR_OUTPUT
	USIALARMGROUPID : ALARMGROUP_ID;
	UIALARMID : ALARM_ID;
END_VAR
END_METHOD

METHOD RAISEEVENTALARMINSTANCE : BOOL
VAR_INPUT
	PFBINSTANCE : POINTER TO BYTE;
	UITEMPLATEALARMID : ALARM_ID;
END_VAR
END_METHOD

METHOD RAISEEVENTALARMINSTANCEBYNAME : BOOL
VAR_INPUT
	PFBINSTANCE : POINTER TO BYTE;
	UITEMPLATEALARMID : ALARM_ID;
	STALARMTEMPLATENAME : STRING(255);
END_VAR
END_METHOD

(* ---- IALARMHANDLER8.itf ---- *)
INTERFACE IALARMHANDLER8
END_INTERFACE

(* ---- IALARMHANDLER9.itf ---- *)
INTERFACE IALARMHANDLER9
END_INTERFACE

METHOD ACTIVATEALARM : BOOL
VAR_INPUT
	USIALARMGROUPID : ALARMGROUP_ID;
	UIALARMID : ALARM_ID;
END_VAR
END_METHOD

METHOD ACTIVATEALARMINSTANCE : BOOL
VAR_INPUT
	PFBINSTANCE : POINTER TO BYTE;
	UITEMPLATEALARMID : ALARM_ID;
END_VAR
END_METHOD

METHOD DEACTIVATEALARM : BOOL
VAR_INPUT
	USIALARMGROUPID : ALARMGROUP_ID;
	UIALARMID : ALARM_ID;
END_VAR
END_METHOD

METHOD DEACTIVATEALARMINSTANCE : BOOL
VAR_INPUT
	PFBINSTANCE : POINTER TO BYTE;
	UITEMPLATEALARMID : ALARM_ID;
END_VAR
END_METHOD

(* ---- IALARMHANDLERREMOTE.itf ---- *)
INTERFACE IALARMHANDLERREMOTE
END_INTERFACE

METHOD GETACTIVEALARMSFROMPROXY
VAR_INPUT
	PASNAME : POINTER TO ARRAY [0..10] OF STRING;
	IGROUPCOUNT : INT;
	FILTERCRITERIA : REFERENCE TO VisuFbAlarmFilterCriteria;
	ITFALARMDATABLOCK : IAlarmDataBlockBaseDINT;
END_VAR
VAR_IN_OUT
	DISTUBPROG : DINT;
END_VAR
END_METHOD

METHOD GETALARMCLASSDESCBYNAMEFROMPROXY
VAR_INPUT
	SPROXYNAME : STRING;
	SCLASSNAME : STRING;
END_VAR
VAR_OUTPUT
	SDESC : ProxyStructAlarmClassDesc;
END_VAR
END_METHOD

METHOD GETALARMCLASSDESCFROMPROXY
VAR_INPUT
	SNAME : STRING;
	UDIID : UDINT;
END_VAR
VAR_OUTPUT
	SDESC : ProxyStructAlarmClassDesc;
END_VAR
END_METHOD

METHOD GETALARMDESCFROMPROXY
VAR_INPUT
	SNAME : STRING;
	UDIALMID : UDINT;
	UDIGRPID : UDINT;
END_VAR
VAR_OUTPUT
	SDESC : ProxyStructAlarmDesc;
END_VAR
END_METHOD

METHOD GETALARMDISPLAYOPTIONSFROMPROXY
VAR_INPUT
	ITFALARMMETAOBJECTSTUB5 : IAlarmMetaObjectStub5;
	REFDISPLAYOPTIONS : REFERENCE TO DisplayOptions;
END_VAR
VAR_OUTPUT
	XVALID : BOOL;
	SCLASSREMAP : STRING;
END_VAR
END_METHOD

METHOD GETALARMGROUPDESCBYNAMEFROMPROXY
VAR_INPUT
	SPROXYNAME : STRING;
	SGRPNAME : STRING;
END_VAR
VAR_OUTPUT
	SDESC : ProxyStructAlarmGroupDesc;
END_VAR
END_METHOD

METHOD GETALARMGROUPDESCFROMPROXY
VAR_INPUT
	SNAME : STRING;
	UDIID : UDINT;
END_VAR
VAR_OUTPUT
	SDESC : ProxyStructAlarmGroupDesc;
END_VAR
END_METHOD

METHOD GETALARMMESSAGEFROMPROXY
VAR_INPUT
	ITFALARMMETAOBJECTSTUB5 : IAlarmMetaObjectStub5;
	IWHICHMESSAGE : INT;
	REFCHARBUFFERSTRING : REFERENCE TO CharBufferString;
	STRINGTYPE : __SYSTEM.TYPE_CLASS;
END_VAR
END_METHOD

METHOD GETALARMMESSAGEFROMPROXY2
VAR_INPUT
	SNAME : STRING;
	STEXTLISTNAME : STRING;
	STEXTLISTINDEX : STRING;
	IWHICHMESSAGE : INT;
	STRINGTYPE : __SYSTEM.TYPE_CLASS;
END_VAR
VAR_OUTPUT
	MESSAGE : CharBufferPtr;
END_VAR
END_METHOD

METHOD GETPROXY : IProxy
VAR_INPUT
	SNAME : STRING;
END_VAR
END_METHOD

METHOD REGISTERALARMCONFIGURATIONREMOTE
VAR_INPUT
	ITFALARMCONFIGURATION : IAlarmConfigurationRemote;
END_VAR
END_METHOD

METHOD SETALARMSTOACKPROXY
VAR_INPUT
	ITFALARMDATABLOCK : IAlarmDataBlockBase2;
END_VAR
END_METHOD

(* ---- IALARMHANDLERREMOTEMONITOR.itf ---- *)
INTERFACE IALARMHANDLERREMOTEMONITOR
END_INTERFACE

METHOD GETPROXYALARMCLASSESDESCRIPTION : BOOL
VAR_INPUT
	SNAME : STRING;
	PCLDESC : POINTER TO ARRAY [0..0] OF ProxyStructMonitorAlarmClassDesc;
	ISIZE : INT;
END_VAR
VAR_OUTPUT
	ICLCNT : INT;
END_VAR
END_METHOD

METHOD GETPROXYALARMGROUPSDESCRIPTION : BOOL
VAR_INPUT
	SNAME : STRING;
	PGRPDESC : POINTER TO ARRAY [0..0] OF ProxyStructMonitorAlarmGroupDesc;
	ISIZE : INT;
END_VAR
VAR_OUTPUT
	IGRPCNT : INT;
END_VAR
END_METHOD

METHOD GETPROXYALARMSDESCRIPTION : BOOL
VAR_INPUT
	SNAME : STRING;
	PALMDESC : POINTER TO ARRAY [0..0] OF ProxyStructMonitorAlarmDesc;
	DISIZE : DINT;
END_VAR
VAR_OUTPUT
	DIALMCNT : DINT;
END_VAR
END_METHOD

METHOD GETPROXYSTATISTICS : BOOL
VAR_INPUT
	SNAME : STRING;
END_VAR
VAR_OUTPUT
	STRUCTMONITOR : ProxyStructMonitor;
END_VAR
END_METHOD

METHOD GETPROXYSTATISTICSSINGLEACTIVITY : BOOL
VAR_INPUT
	SNAME : STRING;
	ITASKID : INT;
END_VAR
VAR_OUTPUT
	STRUCTMONITOR : ProxyStructMonitorRequest;
END_VAR
END_METHOD

(* ---- IALARMMANAGERCLIENT.itf ---- *)
INTERFACE IALARMMANAGERCLIENT
END_INTERFACE

METHOD ACTIVEALARMSCHANGED
END_METHOD

METHOD ALARMSTORAGEMODIFIED
END_METHOD

METHOD GETFILTERCRITERIA : IAlarmFilterCriteria
END_METHOD

(* ---- IALARMMANAGERCLIENT2.itf ---- *)
INTERFACE IALARMMANAGERCLIENT2
END_INTERFACE

METHOD EVENTOCCURRED
VAR_INPUT
	ITFALARM : IAlarm;
END_VAR
END_METHOD

(* ---- IALARMMETAOBJECTSTUBTARGETVISU.itf ---- *)
INTERFACE IALARMMETAOBJECTSTUBTARGETVISU
END_INTERFACE

METHOD GETALARM : POINTER TO Alarm
END_METHOD

METHOD SETALARM
VAR_INPUT
	PALARM : POINTER TO Alarm;
END_VAR
END_METHOD

METHOD SETCURRENTVALUE
VAR_INPUT
	ITFTYPEDVALUECURRENT : ITypedValue;
END_VAR
END_METHOD

(* ---- IALARMNOTIFIABLE.itf ---- *)
INTERFACE IALARMNOTIFIABLE
END_INTERFACE

METHOD EXECUTE
VAR_INPUT
	ECURRTRANSITION : AlarmStateTransition;
	ITFALARM : IAlarm;
	PBYADDITIONALDATA : POINTER TO BYTE;
END_VAR
END_METHOD

(* ---- IALARMOBSERVATIONTYPE.itf ---- *)
INTERFACE IALARMOBSERVATIONTYPE
END_INTERFACE

METHOD ISACTIVE : BOOL
VAR_INPUT
	ECURRSTATE : AlarmState;
END_VAR
END_METHOD

METHOD ISIMMEDIATELYACTIVE : BOOL
END_METHOD

(* ---- IALARMREMOTE.itf ---- *)
INTERFACE IALARMREMOTE
END_INTERFACE

(* ---- IALARMSCALLONINITIALIZE.itf ---- *)
INTERFACE IALARMSCALLONINITIALIZE
END_INTERFACE

(* ---- IALARMSTATECHANGEDEVENTLISTENER.itf ---- *)
INTERFACE IALARMSTATECHANGEDEVENTLISTENER
END_INTERFACE

METHOD ACTIONSTATECHANGED : BOOL
VAR_INPUT
	ITFALARM : IAlarm;
	ESTATEOLD : AlarmState;
	ESTATENEW : AlarmState;
	ESTATETRANSITION : AlarmStateTransition;
END_VAR
END_METHOD

METHOD DEACTIVATIONSTATECHANGED : BOOL
VAR_INPUT
	ITFALARM : IAlarm;
	XNEWDEACTIVATIONSTATE : BOOL;
END_VAR
END_METHOD

METHOD REGISTERLISTENER : BOOL
VAR_INPUT
	ITFALARMSTATECHANGEDLISTENER : IAlarmStateChangedListener;
END_VAR
END_METHOD

(* ---- IALARMSTATECHANGEDLISTENER.itf ---- *)
INTERFACE IALARMSTATECHANGEDLISTENER
END_INTERFACE

METHOD ALARMSTATECHANGED : BOOL
VAR_INPUT
	ITFALARM5 : IAlarm5;
	EOLDSTATE : AlarmState;
	ENEWSTATE : AlarmState;
	ESTATETRANSITION : AlarmStateTransition;
END_VAR
END_METHOD

(* ---- IALARMSTATECHANGEDLISTENER2.itf ---- *)
INTERFACE IALARMSTATECHANGEDLISTENER2
END_INTERFACE

METHOD ALARMDEACTIVATIONSTATECHANGED : BOOL
VAR_INPUT
	ITFALARM5 : IAlarm5;
	XNEWDEACTIVATIONSTATE : BOOL;
END_VAR
END_METHOD

(* ---- IALARMSTATEMACHINE.itf ---- *)
INTERFACE IALARMSTATEMACHINE
END_INTERFACE

METHOD DOACKNOWLEDGE : AlarmState
VAR_INPUT
	ECURRENTSTATE : AlarmState;
END_VAR
VAR_OUTPUT
	ESTATETRANSITION : AlarmStateTransition;
END_VAR
END_METHOD

METHOD DOACTIVATE : AlarmState
VAR_INPUT
	ECURRENTSTATE : AlarmState;
END_VAR
END_METHOD

METHOD DODEACTIVATE : AlarmState
VAR_INPUT
	ECURRENTSTATE : AlarmState;
END_VAR
VAR_OUTPUT
	ESTATETRANSITION : AlarmStateTransition;
END_VAR
END_METHOD

(* ---- IALARMSTORAGEDATACOMPARER.itf ---- *)
INTERFACE IALARMSTORAGEDATACOMPARER
END_INTERFACE

METHOD COMPARE : INT
VAR_INPUT
	DIINDEXALARM1 : DINT;
	DIINDEXALARM2 : DINT;
END_VAR
END_METHOD

METHOD INITIALIZE
VAR_INPUT
	ITFRANDOMALARMREADACCESS : IRandomAlarmReadAccess;
END_VAR
END_METHOD

(* ---- IALARMSTORAGELISTENER.itf ---- *)
INTERFACE IALARMSTORAGELISTENER
END_INTERFACE

METHOD ALARMADDED
VAR_INPUT
	ALARM : AlarmStorageRow;
END_VAR
END_METHOD

METHOD ALARMMODIFIED
VAR_INPUT
	ALARM : AlarmStorageRow;
END_VAR
END_METHOD

(* ---- IALARMSTORAGELISTENER2.itf ---- *)
INTERFACE IALARMSTORAGELISTENER2
END_INTERFACE

METHOD ALARMDELETED
VAR_INPUT
	IDROW : CAA.IDENT;
END_VAR
END_METHOD

(* ---- IALARMSTORAGELISTENER3.itf ---- *)
INTERFACE IALARMSTORAGELISTENER3
END_INTERFACE

METHOD ALARMCLEARFINISHED
END_METHOD

(* ---- IALARMSTORAGEMANAGER.itf ---- *)
INTERFACE IALARMSTORAGEMANAGER
END_INTERFACE

METHOD BEGINTRANSACTION : STO.ITransaction
VAR_INPUT
	XREADONLY : BOOL;
END_VAR
VAR_OUTPUT
	EERROR : STO.ERROR;
END_VAR
END_METHOD

METHOD CLOSETABLE
VAR_INPUT
	ITFTABLE : STO.ITable;
END_VAR
END_METHOD

METHOD DETERMINEROOTPAGES : STO.ERROR
END_METHOD

METHOD ENDTRANSACTION
VAR_INPUT
	ITFTRANSACTION : STO.ITransaction;
	EERROR : STO.ERROR;
END_VAR
END_METHOD

METHOD GETCOLUMNIDENTIFIER : CAA.IDENT
VAR_INPUT
	IDCOLUMN : CAA.IDENT;
END_VAR
END_METHOD

METHOD GETNUMBEROFLATCHVARIABLES : CAA.COUNT
VAR_INPUT
	IDBVERSION : INT;
	UDICOUNTCOLUMNSTBLALARM : CAA.COUNT;
END_VAR
END_METHOD

METHOD GETROOTPAGE : CAA.IDENT
VAR_INPUT
	EDATABASEOBJECT : EAlarmStorageObject;
END_VAR
END_METHOD

METHOD GETSTORAGE : STO.IStorage
END_METHOD

METHOD OPENTABLE : STO.ITable
VAR_INPUT
	XREADONLY : BOOL;
END_VAR
VAR_OUTPUT
	EERROR : STO.ERROR;
END_VAR
END_METHOD

(* ---- IALARMSTORAGEREADERCONSUMER.itf ---- *)
INTERFACE IALARMSTORAGEREADERCONSUMER
END_INTERFACE

METHOD ALARMREAD
VAR_INPUT
	DIWHICHROW : DINT;
	STATICDATA : AlarmStorageStaticData;
END_VAR
END_METHOD

METHOD BEFOREREADING
VAR_INPUT
	USICOUNTLATCHVARIABLES : USINT;
END_VAR
END_METHOD

METHOD LATCHVARIABLEREAD
VAR_INPUT
	DIWHICHROW : DINT;
	USIWHICHVARIABLE : USINT;
	LILATCHVARVALUE : LINT;
	ILATCHVARTYPE : TypeClass;
	XVALUENULL : BOOL;
END_VAR
END_METHOD

METHOD READINGDATACOMPLETED
END_METHOD

(* ---- IALARMSTORAGEREADERCONSUMER2.itf ---- *)
INTERFACE IALARMSTORAGEREADERCONSUMER2
END_INTERFACE

(* ---- IALARMTRAVERSALCONSUMER.itf ---- *)
INTERFACE IALARMTRAVERSALCONSUMER
END_INTERFACE

METHOD AFTERLASTALARMOFALARMGROUP
VAR_INPUT
	ITFALARMGROUP : IAlarmGroup;
END_VAR
END_METHOD

METHOD ALARMCLASSREACHED
VAR_INPUT
	ITFALARMCLASS : IAlarmClass;
END_VAR
END_METHOD

METHOD ALARMHISTORICALISRELEVANT : BOOL
VAR_INPUT
	ROW : REFERENCE TO AlarmStorageRow;
END_VAR
END_METHOD

METHOD ALARMHISTORICALREACHED : UDINT
VAR_INPUT
	ROW : REFERENCE TO AlarmStorageRow;
END_VAR
END_METHOD

METHOD ALARMREACHED
VAR_INPUT
	IWHICHALARMGROUP : INT;
	IWHICHALARM : INT;
	ITFALARM : IAlarm3;
END_VAR
END_METHOD

METHOD BEFOREFIRSTALARMOFALARMGROUP
VAR_INPUT
	ITFALARMGROUP : IAlarmGroup;
END_VAR
END_METHOD

METHOD BEGINTRAVERSAL
END_METHOD

METHOD ENDTRAVERSAL
END_METHOD

METHOD GETACTIVEALARMHISTORICALROWID
VAR_INPUT
	XFIRST : BOOL;
END_VAR
VAR_OUTPUT
	DWROWID : DWORD;
	LITS : LINT;
END_VAR
END_METHOD

(* ---- IALMCONFIGSERVICECONSUMER.itf ---- *)
INTERFACE IALMCONFIGSERVICECONSUMER
END_INTERFACE

(* ---- IALMCONFIGSERVICEPROVIDER.itf ---- *)
INTERFACE IALMCONFIGSERVICEPROVIDER
END_INTERFACE

METHOD GETPROXYALARMCLASSDESCRIPTIONOBJECT : POINTER TO ProxyStructAlarmClass
VAR_INPUT
	IOBJNUM : INT;
END_VAR
END_METHOD

METHOD GETPROXYALARMDESCRIPTIONOBJECT : POINTER TO ProxyStructAlarm
VAR_INPUT
	IOBJNUM : INT;
END_VAR
END_METHOD

METHOD GETPROXYALARMGROUPDESCRIPTIONOBJECT : POINTER TO ProxyStructAlarmGroup
VAR_INPUT
	IOBJNUM : INT;
END_VAR
END_METHOD

(* ---- IALMRECORDSERVICECONSUMER.itf ---- *)
INTERFACE IALMRECORDSERVICECONSUMER
END_INTERFACE

METHOD SETALARMMANAGERLIBVERSION
VAR_INPUT
	LIBVER : VERSION;
END_VAR
END_METHOD

METHOD SETALARMSCOUNT
VAR_INPUT
	DIVALUE : DINT;
END_VAR
END_METHOD

METHOD SETCLASSESCOUNT
VAR_INPUT
	IVALUE : INT;
END_VAR
END_METHOD

METHOD SETRECORDID
VAR_INPUT
	IVALUE : INT;
END_VAR
END_METHOD

(* ---- IALMRECORDSERVICEPROVIDER.itf ---- *)
INTERFACE IALMRECORDSERVICEPROVIDER
END_INTERFACE

METHOD GETALARMGROUP : STRING
VAR_INPUT
	IWHICHALARMGROUP : INT;
END_VAR
END_METHOD

METHOD GETALARMGROUPSNUM : INT
END_METHOD

(* ---- ICHANGEEVALUATOR.itf ---- *)
INTERFACE ICHANGEEVALUATOR
END_INTERFACE

METHOD HASCHANGED : BOOL
VAR_INPUT
	UIID : ALARM_ID;
END_VAR
END_METHOD

(* ---- ICHANNELTESTSERVICECONSUMER.itf ---- *)
INTERFACE ICHANNELTESTSERVICECONSUMER
END_INTERFACE

METHOD SETVALUE
VAR_INPUT
	IVALUE : INT;
END_VAR
END_METHOD

(* ---- ICHANNELTESTSERVICEPROVIDER.itf ---- *)
INTERFACE ICHANNELTESTSERVICEPROVIDER
END_INTERFACE

METHOD GETVALUE : INT
END_METHOD

(* ---- IDATABASEACCESS.itf ---- *)
INTERFACE IDATABASEACCESS
END_INTERFACE

METHOD CALLINGMETHODORFUNCTIONENTER
VAR_INPUT
	ICALLINGMETHOD : INT;
END_VAR
END_METHOD

METHOD CALLINGMETHODORFUNCTIONLEAVE
END_METHOD

METHOD GETNUMBEROFLATCHVARIABLES : USINT
END_METHOD

METHOD GETROOTPAGE : CAA.IDENT
VAR_INPUT
	EWHICHALARMSTORAGEOBJECT : EAlarmStorageObject;
END_VAR
END_METHOD

METHOD ISONLYONEALARMCLASSSELECTED : BOOL
END_METHOD

METHOD ISONLYONEALARMGROUPSELECTED : BOOL
END_METHOD

METHOD PREPAREDATABASEACCESS : STO.ERROR
END_METHOD

METHOD TBLALARMCURSORCLOSE : STO.ERROR
VAR_INPUT
	EERRORFROMPREVIOUSPROCESSING : STO.ERROR;
END_VAR
END_METHOD

METHOD TBLALARMCURSORMOVE : STO.ERROR
VAR_INPUT
	EDIRECTION : STO.DIRECTION;
END_VAR
VAR_OUTPUT
	XEOF : BOOL;
END_VAR
END_METHOD

METHOD TBLALARMCURSOROPEN : STO.ERROR
VAR_INPUT
	FILTERCRITERIA : REFERENCE TO VisuFbAlarmFilterCriteria;
END_VAR
END_METHOD

METHOD TBLALARMCURSOROPEN2 : STO.ERROR
VAR_INPUT
	IDINDEX : CAA.IDENT;
END_VAR
END_METHOD

METHOD TBLALARMCURSORSETPOSITION : STO.ERROR
VAR_INPUT
	FILTERCRITERIA : REFERENCE TO VisuFbAlarmFilterCriteria;
	BROWIDVALID : BOOL;
	DIROWID : DINT;
END_VAR
END_METHOD

METHOD TBLALARMGETLATCHVARTYPE : STO.ERROR
VAR_INPUT
	IDWHICHCOLUMN : CAA.IDENT;
	USIWHICHLATCHVAR : USINT;
END_VAR
VAR_OUTPUT
	BYTYPE : BYTE;
	XNULL : BOOL;
END_VAR
END_METHOD

METHOD TBLALARMGETLATCHVARVALUE : STO.ERROR
VAR_INPUT
	IDWHICHCOLUMN : CAA.IDENT;
	USIWHICHLATCHVAR : USINT;
END_VAR
VAR_OUTPUT
	LIVALUE : LINT;
	XNULL : BOOL;
END_VAR
END_METHOD

METHOD TBLALARMGETMINMAXROWIDS : BOOL
VAR_OUTPUT
	IDROWMIN : LINT;
	IDROWMAX : LINT;
	EERROR : STO.ERROR;
END_VAR
END_METHOD

METHOD TBLALARMGETROWCOUNT : CAA.COUNT
VAR_OUTPUT
	EERROR : STO.ERROR;
END_VAR
END_METHOD

METHOD TBLALARMGETTIMESTAMPVALUE : LINT
VAR_INPUT
	IDWHICHCOLUMN : CAA.IDENT;
END_VAR
VAR_OUTPUT
	EERROR : STO.ERROR;
END_VAR
END_METHOD

METHOD TBLALARMGET_DINT : STO.ERROR
VAR_INPUT
	IDWHICHCOLUMN : CAA.IDENT;
	IWHICHCOLUMN : INT;
END_VAR
VAR_OUTPUT
	DIVALUE : DINT;
	XNULL : BOOL;
END_VAR
END_METHOD

METHOD TBLALARMGET_LINT : STO.ERROR
VAR_INPUT
	IDWHICHCOLUMN : CAA.IDENT;
	IWHICHCOLUMN : INT;
END_VAR
VAR_OUTPUT
	LIVALUE : LINT;
	XNULL : BOOL;
END_VAR
END_METHOD

METHOD TBLALARMGET_SINT : STO.ERROR
VAR_INPUT
	IDWHICHCOLUMN : CAA.IDENT;
	IWHICHCOLUMN : INT;
END_VAR
VAR_OUTPUT
	SIVALUE : SINT;
	XNULL : BOOL;
END_VAR
END_METHOD

METHOD TBLALARMISNOTEMPTY : BOOL
VAR_OUTPUT
	EERROR : STO.ERROR;
END_VAR
END_METHOD

METHOD TBLALARMROWGETCURRENT : STO.ERROR
END_METHOD

METHOD TBLALARMROWGETCURRENTID : DINT
END_METHOD

METHOD TBLALARMROWISVALID : BOOL
END_METHOD

METHOD TBLALARMROWRELEASE : STO.ERROR
VAR_INPUT
	EERRORFROMPREVIOUSPROCESSING : STO.ERROR;
END_VAR
END_METHOD

METHOD TBLALARMROWSELECT : STO.ERROR
VAR_INPUT
	IDROW : CAA.IDENT;
	XDOERRORHANDLING : BOOL;
END_VAR
END_METHOD

METHOD TBLALARMTABLECLOSE : STO.ERROR
END_METHOD

METHOD TBLALARMTABLEISOPEN : BOOL
END_METHOD

METHOD TBLALARMTABLEOPEN : STO.ERROR
VAR_INPUT
	XREADONLY : BOOL;
END_VAR
END_METHOD

METHOD TBLLATCHVARSTRINGSCLOSEIFNEEDED : STO.ERROR
VAR_INPUT
	EERRORFROMPREVIOUSPROCESSING : STO.ERROR;
END_VAR
END_METHOD

METHOD TBLLATCHVARSTRINGSCURSORSEARCHROWID : STO.ERROR
VAR_INPUT
	LIROWID : LINT;
END_VAR
END_METHOD

METHOD TBLLATCHVARSTRINGSGET_TEXT : STO.ERROR
VAR_INPUT
	IDWHICHCOLUMN : CAA.IDENT;
	IWHICHCOLUMN : INT;
END_VAR
VAR_OUTPUT
	XNULL : BOOL;
END_VAR
VAR_IN_OUT
	TXTVALUE : STO.TEXT;
END_VAR
END_METHOD

METHOD TBLLATCHVARSTRINGSOPENIFNEEDED : STO.ERROR
END_METHOD

METHOD TBLLATCHVARSTRINGSROWGETCURRENT : STO.ERROR
END_METHOD

METHOD TBLLATCHVARSTRINGSROWRELEASE : STO.ERROR
VAR_INPUT
	EERRORFROMPREVIOUSPROCESSING : STO.ERROR;
END_VAR
END_METHOD

METHOD TEXTCOPYTOSTRING : STO.ERROR
VAR_INPUT
	XFREE : BOOL;
END_VAR
VAR_IN_OUT
	TXTVALUE : STO.TEXT;
	SVALUE : STRING(1);
	SZVALUE : CAA.SIZE;
END_VAR
END_METHOD

METHOD TEXTCOPYTOWSTRING : STO.ERROR
VAR_INPUT
	XFREE : BOOL;
END_VAR
VAR_IN_OUT
	TXTVALUE : STO.TEXT;
	WSVALUE : WSTRING(1);
	SZVALUE : CAA.SIZE;
END_VAR
END_METHOD

METHOD TRANSACTIONBEGIN : STO.ERROR
VAR_INPUT
	XREADONLY : BOOL;
END_VAR
END_METHOD

METHOD TRANSACTIONBEGINFAILED : BOOL
END_METHOD

METHOD TRANSACTIONEND
VAR_INPUT
	EERRORFROMPREVIOUSPROCESSING : STO.ERROR;
END_VAR
END_METHOD

(* ---- IDATABASEACCESS2.itf ---- *)
INTERFACE IDATABASEACCESS2
END_INTERFACE

METHOD TBLALARMGET_INT : STO.ERROR
VAR_INPUT
	IDWHICHCOLUMN : CAA.IDENT;
	IWHICHCOLUMN : INT;
END_VAR
VAR_OUTPUT
	IVALUE : INT;
	XNULL : BOOL;
END_VAR
END_METHOD

METHOD TBLVERSIONGETCURRENT : STO.ERROR
VAR_OUTPUT
	IVERSION : INT;
END_VAR
END_METHOD

(* ---- IDATABASEACCESS3.itf ---- *)
INTERFACE IDATABASEACCESS3
END_INTERFACE

METHOD GETRELEVANTFILTERDATA
VAR_OUTPUT
	EDBBYTEORDER : EAlarmByteOrder;
END_VAR
END_METHOD

METHOD TBLALARMCURSORSEARCHROWID : STO.ERROR
VAR_INPUT
	IDROW : DINT;
END_VAR
END_METHOD

METHOD TBLGETBYTEORDER : STO.ERROR
VAR_OUTPUT
	EBYTEORDER : EAlarmByteOrder;
END_VAR
END_METHOD

METHOD TBLVERSIONGETCURRENT2 : STO.ERROR
VAR_OUTPUT
	IVERSION : INT;
	EDBUSED : EDBType;
END_VAR
END_METHOD

(* ---- IDATABASEACCESS4.itf ---- *)
INTERFACE IDATABASEACCESS4
END_INTERFACE

METHOD TBLALARMGETCOMMENTVALUE : STO.ERROR
VAR_INPUT
	IDWHICHCOLUMN : CAA.IDENT;
	IWHICHCOLUMN : INT;
END_VAR
VAR_OUTPUT
	XNULL : BOOL;
END_VAR
VAR_IN_OUT
	WSVALUE : WSTRING(2000);
END_VAR
END_METHOD

(* ---- IDATABASEFILEALARMSTORAGE.itf ---- *)
INTERFACE IDATABASEFILEALARMSTORAGE
END_INTERFACE

METHOD CLOSETABLE
VAR_INPUT
	ITFTABLE : STO.ITable;
END_VAR
END_METHOD

METHOD GETDATABASEFILEPATH : STRING
END_METHOD

METHOD GETFILELIMIT : FileLimit
END_METHOD

METHOD GETMAXRECORDCOUNT : UDINT
END_METHOD

METHOD GETSUBDIRECTORY : STRING
END_METHOD

METHOD OPENTABLE : STO.ITable
VAR_INPUT
	XREADONLY : BOOL;
END_VAR
VAR_OUTPUT
	EERROR : STO.ERROR;
END_VAR
END_METHOD

METHOD WRITETOSTORAGE : STO.ERROR
VAR_INPUT
	ITFTABLE : STO.ITable;
	ROW : AlarmStorageRow;
	ICOUNTRETRIES : INT;
END_VAR
END_METHOD

(* ---- IDATABASEFILEALARMSTORAGE10.itf ---- *)
INTERFACE IDATABASEFILEALARMSTORAGE10
END_INTERFACE

(* ---- IDATABASEFILEALARMSTORAGE11.itf ---- *)
INTERFACE IDATABASEFILEALARMSTORAGE11
END_INTERFACE

METHOD CLEARBUFFER
END_METHOD

(* ---- IDATABASEFILEALARMSTORAGE2.itf ---- *)
INTERFACE IDATABASEFILEALARMSTORAGE2
END_INTERFACE

METHOD ADDALARMSTORAGELISTENER : EAlarmStorageReaderErrors
VAR_INPUT
	ITFALARMSTORAGELISTENER : IAlarmStorageListener;
END_VAR
END_METHOD

METHOD CREATEALARMSTORAGEMETADATAFILE
VAR_INPUT
	UDICOUNTCOLUMNSTBLALARM : CAA.COUNT;
END_VAR
END_METHOD

METHOD OPENTABLE2 : STO.ITable
VAR_INPUT
	XREADONLY : BOOL;
END_VAR
VAR_OUTPUT
	EERROR : STO.ERROR;
END_VAR
END_METHOD

METHOD REMOVEALARMSTORAGELISTENER : EAlarmStorageReaderErrors
VAR_INPUT
	ITFALARMSTORAGELISTENER : IAlarmStorageListener;
END_VAR
END_METHOD

(* ---- IDATABASEFILEALARMSTORAGE3.itf ---- *)
INTERFACE IDATABASEFILEALARMSTORAGE3
END_INTERFACE

METHOD CHECKFILELIMITREACHED : STO.Error
VAR_INPUT
	ITFTABLE : STO.ITable;
	ICOUNTRETRIES : INT;
	ICOUNTROWSTOINSERT : INT;
END_VAR
END_METHOD

METHOD ENDTRANSACTION
VAR_INPUT
	ITFTRANSACTION : STO.ITransaction;
	EERROR : STO.ERROR;
END_VAR
END_METHOD

METHOD GETEXCLUSIVETRANSACTION : STO.ITransaction
VAR_INPUT
	ICOUNTRETRIES : INT;
END_VAR
VAR_OUTPUT
	EERROR : STO.ERROR;
END_VAR
END_METHOD

METHOD WRITETOSTORAGE2 : STO.ERROR
VAR_INPUT
	ITFTABLE : STO.ITable;
	ROW : AlarmStorageRow;
	ITFTRANSACTION : STO.ITransaction;
END_VAR
END_METHOD

(* ---- IDATABASEFILEALARMSTORAGE4.itf ---- *)
INTERFACE IDATABASEFILEALARMSTORAGE4
END_INTERFACE

METHOD DELETEALARMSTORAGEFILE : STO.ERROR
VAR_INPUT
	SFILEPATH : CAA.FILENAME;
END_VAR
END_METHOD

METHOD GETALARMSFROMSTORAGE : STO.ERROR
VAR_INPUT
	ISKIPROWS : INT;
	IMAXROWS : INT;
	FILTERCRITERIA : REFERENCE TO VisuFbAlarmFilterCriteria;
	ITFALARMDATABLOCK : IAlarmDataBlockBase2;
END_VAR
VAR_IN_OUT
	BROWIDVALID : BOOL;
	DIROWID : DINT;
END_VAR
END_METHOD

METHOD GETCOUNTALARMSFROMSTORAGE : DINT
VAR_INPUT
	FILTERCRITERIA : REFERENCE TO VisuFbAlarmFilterCriteria;
	ITFALARMDATABLOCK : IAlarmDataBlockBase2;
END_VAR
VAR_OUTPUT
	EERROR : STO.ERROR;
	DWCOUNTLATCHVARIABLESINSTORAGE : CAA.COUNT;
END_VAR
END_METHOD

(* ---- IDATABASEFILEALARMSTORAGE5.itf ---- *)
INTERFACE IDATABASEFILEALARMSTORAGE5
END_INTERFACE

METHOD CREATEWRITECONTEXT : IDatabaseFileWriteContext
END_METHOD

METHOD SCANSTORAGE : STO.ERROR
VAR_INPUT
	ITFCONSUMER : IRemoteDeviceTraversalConsumer;
END_VAR
VAR_OUTPUT
	IVERSION : INT;
	DIREMOTEENTRIESCNT : DINT;
END_VAR
END_METHOD

METHOD WRITETOSTORAGE3 : STO.ERROR
VAR_INPUT
	WRITECONTEXT : IDatabaseFileWriteContext;
	ROW : AlarmStorageRow;
	XFORCEINSERT : BOOL;
	XFIRST : BOOL;
END_VAR
END_METHOD

(* ---- IDATABASEFILEALARMSTORAGE6.itf ---- *)
INTERFACE IDATABASEFILEALARMSTORAGE6
END_INTERFACE

METHOD CLEARALARMSINSTATENORMAL : STO.Error
VAR_INPUT
	ITFTABLE : STO.ITable;
END_VAR
VAR_OUTPUT
	XFINISHED : BOOL;
END_VAR
VAR_IN_OUT
	DIREMAININGROWCOUNT : DINT;
END_VAR
END_METHOD

METHOD ROWSELECT : STO.IRow
VAR_INPUT
	ITFTABLE : STO.ITable;
	IDROW : CAA.IDENT;
END_VAR
END_METHOD

(* ---- IDATABASEFILEALARMSTORAGE7.itf ---- *)
INTERFACE IDATABASEFILEALARMSTORAGE7
END_INTERFACE

METHOD CHECKRECORDLIMITREACHED : STO.Error
VAR_INPUT
	ITFTABLE : STO.ITable;
	ICOUNTRETRIES : INT;
	ICOUNTROWSTOINSERT : INT;
	XFORCE : BOOL;
END_VAR
VAR_OUTPUT
	XLIMIT : BOOL;
	UDIMAXRECORDCOUNT : UDINT;
END_VAR
END_METHOD

METHOD DELETEALARMS : STO.Error
VAR_INPUT
	ITFTABLE : STO.ITable;
	ICOUNTRETRIES : INT;
	DICOUNTROWSTODELETE : DINT;
END_VAR
VAR_OUTPUT
	DIROWSDELETED : DINT;
END_VAR
END_METHOD

METHOD GETRECORDSIZE : INT
END_METHOD

METHOD GETSTORAGESIZE : LINT
END_METHOD

(* ---- IDATABASEFILEALARMSTORAGE8.itf ---- *)
INTERFACE IDATABASEFILEALARMSTORAGE8
END_INTERFACE

METHOD SETEMPTYTIMESTAMPINACTIVETOSTARTTIME : STO.Error
VAR_INPUT
	ITFTABLE : STO.ITable;
END_VAR
END_METHOD

(* ---- IDATABASEFILEALARMSTORAGE9.itf ---- *)
INTERFACE IDATABASEFILEALARMSTORAGE9
END_INTERFACE

METHOD CHECKFILELIMITREACHEDUDINT : STO.Error
VAR_INPUT
	ITFTABLE : STO.ITable;
	ICOUNTRETRIES : INT;
	UDICOUNTROWSTOINSERT : UDINT;
END_VAR
END_METHOD

METHOD CHECKRECORDLIMITREACHEDUDINT : STO.Error
VAR_INPUT
	ITFTABLE : STO.ITable;
	ICOUNTRETRIES : INT;
	UDICOUNTROWSTOINSERT : UDINT;
	XFORCE : BOOL;
END_VAR
VAR_OUTPUT
	XLIMIT : BOOL;
	UDIMAXRECORDCOUNT : UDINT;
END_VAR
END_METHOD

(* ---- IDATABASEFILEWRITECONTEXT.itf ---- *)
INTERFACE IDATABASEFILEWRITECONTEXT
END_INTERFACE

METHOD GETSTRINGLATCHTABLE : STO.ITable
VAR_OUTPUT
	EERROR : STO.ERROR;
END_VAR
END_METHOD

METHOD RELEASE
VAR_INPUT
	EERRORFORCOMMIT : STO.ERROR;
END_VAR
END_METHOD

(* ---- IDATABASESIZELIMIT.itf ---- *)
INTERFACE IDATABASESIZELIMIT
END_INTERFACE

(* ---- IDEACTIVATOR.itf ---- *)
INTERFACE IDEACTIVATOR
END_INTERFACE

METHOD ISDEACTIVATED : BOOL
VAR_INPUT
	UIID : ALARM_ID;
END_VAR
END_METHOD

(* ---- IEXPRESSIONEVALUATOR.itf ---- *)
INTERFACE IEXPRESSIONEVALUATOR
END_INTERFACE

METHOD ISTRUE : BOOL
VAR_INPUT
	UIID : ALARM_ID;
	ECURRSTATE : AlarmState;
END_VAR
END_METHOD

(* ---- IHASHTABLEKEYELEMENT.itf ---- *)
INTERFACE IHASHTABLEKEYELEMENT
END_INTERFACE

(* ---- IHASHTABLEVALUEELEMENT.itf ---- *)
INTERFACE IHASHTABLEVALUEELEMENT
END_INTERFACE

(* ---- IHISTORICALMSERVICECONSUMER.itf ---- *)
INTERFACE IHISTORICALMSERVICECONSUMER
END_INTERFACE

METHOD SETHASSTORAGE
VAR_INPUT
	XVALUE : BOOL;
END_VAR
END_METHOD

METHOD SETHISTACTIVEALARMSREAD
VAR_INPUT
	ICOUNT : INT;
END_VAR
END_METHOD

METHOD SETHISTALARMSREAD
VAR_INPUT
	DWROWIDLAST : DWORD;
	ICOUNT : INT;
	DISTORAGEROWSCOUNT : DINT;
	ISTORAGECLEAR : INT;
END_VAR
END_METHOD

METHOD SETROWIDS
VAR_INPUT
	DWROWIDFIRST : DWORD;
	DWROWIDLAST : DWORD;
END_VAR
END_METHOD

(* ---- IHISTORICALMSERVICEPROVIDER.itf ---- *)
INTERFACE IHISTORICALMSERVICEPROVIDER
END_INTERFACE

METHOD GETPROXYHISTORICALALARMOBJECT : POINTER TO ProxyFbAlarmHistorical
VAR_INPUT
	XACTIVE : BOOL;
	IOBJNUM : INT;
END_VAR
END_METHOD

METHOD GETRECORDIDHISTORICAL : INT
END_METHOD

METHOD GETROWIDHISTORICALACTIVEALARMS
VAR_INPUT
	XFIRSTCALL : BOOL;
END_VAR
VAR_OUTPUT
	DWROWID : DWORD;
	LITS : LINT;
END_VAR
END_METHOD

METHOD GETROWTOREAD
VAR_OUTPUT
	DWROWIDLAST : DWORD;
	IROWCOUNT : INT;
END_VAR
END_METHOD

(* ---- ILISTELEMENT.itf ---- *)
INTERFACE ILISTELEMENT
END_INTERFACE

METHOD GETLATCHVARIABLES : BOOL
VAR_OUTPUT
	PALATCHVARIABLES : POINTER TO ARRAY [0..255] OF ValueTypeBundle;
	USICOUNTLATCHVARIABLES : USINT;
END_VAR
END_METHOD

METHOD SETLATCHVARIABLES : BOOL
VAR_INPUT
	PALARM : POINTER TO Alarm;
END_VAR
END_METHOD

(* ---- IPROXY.itf ---- *)
INTERFACE IPROXY
END_INTERFACE

METHOD CYCLICCALL : BOOL
END_METHOD

METHOD GETACTIVEALARMS : INT
VAR_INPUT
	SNAME : STRING;
	FILTERCRITERIA : REFERENCE TO VisuFbAlarmFilterCriteria;
	ITFALARMDATABLOCK : IAlarmDataBlockBaseDINT;
END_VAR
VAR_IN_OUT
	DISTUBPROG : DINT;
END_VAR
END_METHOD

METHOD GETACTIVEALARMS2
VAR_INPUT
	FILTERCRITERIA : REFERENCE TO VisuFbAlarmFilterCriteria;
	PAITFALARMS : POINTER TO ARRAY [0..10] OF IAlarm;
	DIARRSIZE : DINT;
END_VAR
VAR_OUTPUT
	DICOUNT : DINT;
END_VAR
END_METHOD

METHOD GETALARMCLASSDESC
VAR_INPUT
	UDIID : UDINT;
END_VAR
VAR_OUTPUT
	SDESC : ProxyStructAlarmClassDesc;
END_VAR
END_METHOD

METHOD GETALARMCLASSDESCBYNAME
VAR_INPUT
	SCLASSNAME : STRING;
END_VAR
VAR_OUTPUT
	SDESC : ProxyStructAlarmClassDesc;
END_VAR
END_METHOD

METHOD GETALARMDESC
VAR_INPUT
	UDIALMID : UDINT;
	UDIGRPID : UDINT;
END_VAR
VAR_OUTPUT
	SDESC : ProxyStructAlarmDesc;
END_VAR
END_METHOD

METHOD GETALARMDISPLAYOPTIONS
VAR_INPUT
	ITFALARMMETAOBJECTSTUB5 : IAlarmMetaObjectStub5;
	REFDISPLAYOPTIONS : REFERENCE TO DisplayOptions;
END_VAR
VAR_OUTPUT
	XVALID : BOOL;
	SCLASSREMAP : STRING;
END_VAR
END_METHOD

METHOD GETALARMGROUPDESC
VAR_INPUT
	UDIID : UDINT;
END_VAR
VAR_OUTPUT
	SDESC : ProxyStructAlarmGroupDesc;
END_VAR
END_METHOD

METHOD GETALARMGROUPDESCBYNAME
VAR_INPUT
	SGRPNAME : STRING;
END_VAR
VAR_OUTPUT
	SDESC : ProxyStructAlarmGroupDesc;
END_VAR
END_METHOD

METHOD GETALARMMESSAGE
VAR_INPUT
	ITFALARMMETAOBJECTSTUB5 : IAlarmMetaObjectStub5;
	IWHICHMESSAGE : INT;
	REFCHARBUFFERSTRING : REFERENCE TO CharBufferString;
	STRINGTYPE : __SYSTEM.TYPE_CLASS;
END_VAR
END_METHOD

METHOD GETALARMMESSAGE2 : Stu.CharBufferPtr
VAR_INPUT
	STEXTLISTNAME : STRING;
	STEXTLISTINDEX : STRING;
	IWHICHMESSAGE : INT;
	STRINGTYPE : __SYSTEM.TYPE_CLASS;
END_VAR
END_METHOD

METHOD GETPROXYNAME : POINTER TO STRING
END_METHOD

METHOD GETTOTALALARMSCOUNT : DINT
END_METHOD

METHOD INITIALIZE : BOOL
VAR_INPUT
	PPARAM : POINTER TO ProxyStructInitialize;
	ITEST : INT;
END_VAR
END_METHOD

METHOD REGISTERUSERCLIENT
END_METHOD

METHOD SETALARMSTOACK
VAR_INPUT
	ITFALARMMETAOBJECTSTUB : IAlarmMetaObjectStub5;
END_VAR
END_METHOD

METHOD SETINITIALDATAFROMDB
VAR_INPUT
	ROW : REFERENCE TO AlarmStorageRow;
	XFIRST : BOOL;
	IVERSION : INT;
END_VAR
END_METHOD

METHOD SETPARAMS
VAR_INPUT
	PPARAM : POINTER TO ProxyStructParam;
END_VAR
END_METHOD

(* ---- IPROXYALARMOBJECT.itf ---- *)
INTERFACE IPROXYALARMOBJECT
END_INTERFACE

METHOD SETCOUNTLATCHVARIABLES
VAR_INPUT
	USICOUNT : USINT;
END_VAR
END_METHOD

(* ---- IPROXYCOMMCHANNEL.itf ---- *)
INTERFACE IPROXYCOMMCHANNEL
END_INTERFACE

METHOD ADDERROR
VAR_INPUT
	ITASKID : INT;
	UDIERROR : UDINT;
	SMSG : STRING;
END_VAR
END_METHOD

METHOD CLEANSTATISTICS : BOOL
VAR_INPUT
	ITASKID : INT;
END_VAR
END_METHOD

METHOD CYCLICCALL
END_METHOD

METHOD EXECUTEREQUEST : UDINT
VAR_INPUT
	ITASKID : INT;
	XLOCK : BOOL;
	HLOCK : RTS_IEC_HANDLE;
END_VAR
END_METHOD

METHOD GETALARMMESSAGETEXT : BOOL
VAR_INPUT
	ITFALARMMETAOBJECTSTUB5 : IAlarmMetaObjectStub5;
	IWHICHMESSAGE : INT;
	STRINGTYPE : __SYSTEM.TYPE_CLASS;
END_VAR
VAR_OUTPUT
	CBPMESSAGE : CharBufferPtr;
END_VAR
END_METHOD

METHOD GETALARMMESSAGETEXT2 : BOOL
VAR_INPUT
	STEXTLISTNAME : STRING;
	STEXTLISTINDEX : STRING;
	IWHICHMESSAGE : INT;
	STRINGTYPE : __SYSTEM.TYPE_CLASS;
END_VAR
VAR_OUTPUT
	CBPMESSAGE : CharBufferPtr;
END_VAR
END_METHOD

METHOD GETSTATISTICSSINGLEREQ : ProxyStructMonitorRequest
VAR_INPUT
	ITASKID : INT;
END_VAR
END_METHOD

METHOD INITIALIZE
VAR_INPUT
	ITFPROXYCONSUMER : IProxyConsumer;
	ITFPROXYPROVIDER : IProxyProvider;
	IMAXALMGROUPS : INT;
END_VAR
END_METHOD

METHOD ISCHANNELAVAILABLE : BOOL
END_METHOD

METHOD ISREQUESTEXECUTABLE : BOOL
VAR_INPUT
	ITASKID : INT;
	XTRYTOFORCE : BOOL;
END_VAR
END_METHOD

METHOD RESTART
END_METHOD

(* ---- IPROXYCONSUMER.itf ---- *)
INTERFACE IPROXYCONSUMER
END_INTERFACE

METHOD COMMUNICATIONFINISHED
VAR_INPUT
	IREQUESTID : INT;
	XWITHERRORS : BOOL;
END_VAR
END_METHOD

METHOD PROXYMANAGERLOG
VAR_INPUT
	SVAL1 : STRING(255);
	SVAL2 : STRING(255);
	SVAL3 : STRING(255);
	UDISEV : UDINT;
END_VAR
END_METHOD

METHOD SETACTIVEALARMSCOUNT
VAR_INPUT
	DICOUNT : DINT;
END_VAR
END_METHOD

METHOD SETALARMMANAGERLIBVERSION
VAR_INPUT
	LIBVER : VERSION;
END_VAR
END_METHOD

METHOD SETDEVICENAME
VAR_INPUT
	SNAME : STRING;
END_VAR
END_METHOD

METHOD SETHASSTORAGE
VAR_INPUT
	XVALUE : BOOL;
END_VAR
END_METHOD

METHOD SETHISTACTIVEALARMSREAD
VAR_INPUT
	ICOUNT : INT;
END_VAR
END_METHOD

METHOD SETHISTALARMSREAD
VAR_INPUT
	DWROWIDLAST : DWORD;
	ICOUNT : INT;
	DISTORAGEROWSCOUNT : DINT;
	ISTORAGECLEAR : INT;
END_VAR
END_METHOD

METHOD SETLATCHVARSCOUNT
VAR_INPUT
	ICOUNT : INT;
END_VAR
END_METHOD

METHOD SETRECORDID
VAR_INPUT
	IVALUE : INT;
END_VAR
END_METHOD

METHOD SETROWIDS
VAR_INPUT
	DWROWIDFIRST : DWORD;
	DWROWIDLAST : DWORD;
END_VAR
END_METHOD

METHOD SETTOTALALARMSCOUNT
VAR_INPUT
	DICOUNT : DINT;
END_VAR
END_METHOD

METHOD SETTOTALCLASSESCOUNT
VAR_INPUT
	ICOUNT : INT;
END_VAR
END_METHOD

(* ---- IPROXYMONITOR.itf ---- *)
INTERFACE IPROXYMONITOR
END_INTERFACE

METHOD GETALARMCLASSESDESCRIPTION
VAR_INPUT
	PCLDESC : POINTER TO ARRAY [0..0] OF ProxyStructMonitorAlarmClassDesc;
	ISIZE : INT;
END_VAR
VAR_OUTPUT
	ICLCNT : INT;
END_VAR
END_METHOD

METHOD GETALARMGROUPSDESCRIPTION
VAR_INPUT
	PGRPDESC : POINTER TO ARRAY [0..0] OF ProxyStructMonitorAlarmGroupDesc;
	ISIZE : INT;
END_VAR
VAR_OUTPUT
	IGRPCNT : INT;
END_VAR
END_METHOD

METHOD GETALARMSDESCRIPTION
VAR_INPUT
	PALMDESC : POINTER TO ARRAY [0..0] OF ProxyStructMonitorAlarmDesc;
	DISIZE : DINT;
END_VAR
VAR_OUTPUT
	DIALMCNT : DINT;
END_VAR
END_METHOD

METHOD GETSTATISTICS : ProxyStructMonitor
VAR_INPUT
	IRECORD : INT;
END_VAR
END_METHOD

METHOD GETSTATISTICSSINGLEREQ : ProxyStructMonitorRequest
VAR_INPUT
	ITASKID : INT;
END_VAR
END_METHOD

(* ---- IPROXYPROVIDER.itf ---- *)
INTERFACE IPROXYPROVIDER
END_INTERFACE

METHOD GETALARMGROUP : STRING
VAR_INPUT
	IWHICHALARMGROUP : INT;
END_VAR
END_METHOD

METHOD GETALARMGROUPSNUM : INT
END_METHOD

METHOD GETAPPLICATION : STRING
END_METHOD

METHOD GETCOUNTALARMSTOACKNOWLEDGE : INT
END_METHOD

METHOD GETNEXTALARMTOACKNOWLEDGE : BOOL
VAR_INPUT
	XFISRTENTRY : BOOL;
END_VAR
VAR_OUTPUT
	ALARMTOACKNOWLEDGE : AlarmToAcknowledge;
END_VAR
END_METHOD

METHOD GETPROXYACTIVEALARMOBJECT : IProxyAlarmObject
VAR_INPUT
	DIOBJNUM : DINT;
END_VAR
END_METHOD

METHOD GETPROXYALARMCLASSDESCRIPTIONOBJECT : POINTER TO ProxyStructAlarmClass
VAR_INPUT
	IOBJNUM : INT;
END_VAR
END_METHOD

METHOD GETPROXYALARMDESCRIPTIONOBJECT : POINTER TO ProxyStructAlarm
VAR_INPUT
	IOBJNUM : INT;
END_VAR
END_METHOD

METHOD GETPROXYALARMGROUPDESCRIPTIONOBJECT : POINTER TO ProxyStructAlarmGroup
VAR_INPUT
	IOBJNUM : INT;
END_VAR
END_METHOD

METHOD GETPROXYHISTORICALALARMOBJECT : POINTER TO ProxyFbAlarmHistorical
VAR_INPUT
	XACTIVE : BOOL;
	IOBJNUM : INT;
END_VAR
END_METHOD

METHOD GETRECORDID : INT
END_METHOD

METHOD GETRECORDIDHISTORICAL : INT
END_METHOD

METHOD GETROWIDHISTORICALACTIVEALARMS
VAR_INPUT
	XFIRSTCALL : BOOL;
END_VAR
VAR_OUTPUT
	DWROWID : DWORD;
	LITS : LINT;
END_VAR
END_METHOD

METHOD GETROWTOREAD
VAR_OUTPUT
	DWROWIDLAST : DWORD;
	IROWCOUNT : INT;
END_VAR
END_METHOD

(* ---- IRANDOMALARMREADACCESS.itf ---- *)
INTERFACE IRANDOMALARMREADACCESS
END_INTERFACE

METHOD GETALARMCLASSID : BOOL
VAR_INPUT
	DIINDEXALARM : DINT;
END_VAR
VAR_OUTPUT
	UDIALARMCLASSID : UDINT;
END_VAR
END_METHOD

METHOD GETALARMGROUPID : BOOL
VAR_INPUT
	DIINDEXALARM : DINT;
END_VAR
VAR_OUTPUT
	UDIALARMGROUPID : UDINT;
END_VAR
END_METHOD

METHOD GETALARMID : BOOL
VAR_INPUT
	DIINDEXALARM : DINT;
END_VAR
VAR_OUTPUT
	UDIALARMID : UDINT;
END_VAR
END_METHOD

METHOD GETLATCHVARTYPE : BOOL
VAR_INPUT
	DIINDEXALARM : DINT;
	IWHICHLATCHVARIABLE : INT;
END_VAR
VAR_OUTPUT
	BYTYPE : BYTE;
END_VAR
END_METHOD

METHOD GETLATCHVARVALUE : BOOL
VAR_INPUT
	DIINDEXALARM : DINT;
	IWHICHLATCHVARIABLE : INT;
END_VAR
VAR_OUTPUT
	LIVALUE : LINT;
END_VAR
END_METHOD

METHOD GETPRIORITY : BOOL
VAR_INPUT
	DIINDEXALARM : DINT;
END_VAR
VAR_OUTPUT
	USIPRIORITY : USINT;
END_VAR
END_METHOD

METHOD GETROWID : BOOL
VAR_INPUT
	DIINDEXALARM : DINT;
END_VAR
VAR_OUTPUT
	DIROWID : DINT;
END_VAR
END_METHOD

METHOD GETSTATE : BOOL
VAR_INPUT
	DIINDEXALARM : DINT;
END_VAR
VAR_OUTPUT
	BYSTATE : BYTE;
END_VAR
END_METHOD

METHOD GETTSACK : BOOL
VAR_INPUT
	DIINDEXALARM : DINT;
END_VAR
VAR_OUTPUT
	LITIMESTAMP : TIMESTAMP;
END_VAR
END_METHOD

METHOD GETTSACTIVE : BOOL
VAR_INPUT
	DIINDEXALARM : DINT;
END_VAR
VAR_OUTPUT
	LITIMESTAMP : TIMESTAMP;
END_VAR
END_METHOD

METHOD GETTSINACTIVE : BOOL
VAR_INPUT
	DIINDEXALARM : DINT;
END_VAR
VAR_OUTPUT
	LITIMESTAMP : TIMESTAMP;
END_VAR
END_METHOD

METHOD GETTSLAST : BOOL
VAR_INPUT
	DIINDEXALARM : DINT;
END_VAR
VAR_OUTPUT
	LITIMESTAMP : TIMESTAMP;
END_VAR
END_METHOD

METHOD GETTRIGGERVALUE : BOOL
VAR_INPUT
	DIINDEXALARM : DINT;
END_VAR
VAR_OUTPUT
	LIVALUE : LINT;
END_VAR
END_METHOD

METHOD GETTRIGGERVALUETYPE : BOOL
VAR_INPUT
	DIINDEXALARM : DINT;
END_VAR
VAR_OUTPUT
	BYTYPE : BYTE;
END_VAR
END_METHOD

(* ---- IRANDOMALARMREADACCESS2.itf ---- *)
INTERFACE IRANDOMALARMREADACCESS2
END_INTERFACE

METHOD GETREMOTEDEVICENAME : BOOL
VAR_INPUT
	DIINDEXALARM : DINT;
END_VAR
VAR_OUTPUT
	SNAME : STRING(255);
END_VAR
END_METHOD

(* ---- IRANDOMALARMREADACCESS3.itf ---- *)
INTERFACE IRANDOMALARMREADACCESS3
END_INTERFACE

METHOD GETCOMMENT : BOOL
VAR_INPUT
	DIINDEXALARM : DINT;
END_VAR
VAR_OUTPUT
	WSCOMMENT : WSTRING(255);
END_VAR
END_METHOD

METHOD GETUSERID : BOOL
VAR_INPUT
	DIINDEXALARM : DINT;
END_VAR
VAR_OUTPUT
	WSUSERID : WSTRING(255);
END_VAR
END_METHOD

(* ---- IREADACTIVEALARMSSERVICECONSUMER.itf ---- *)
INTERFACE IREADACTIVEALARMSSERVICECONSUMER
END_INTERFACE

METHOD SETACTIVEALARMSCOUNT
VAR_INPUT
	DICOUNT : DINT;
END_VAR
END_METHOD

(* ---- IREADACTIVEALARMSSERVICEPROVIDER.itf ---- *)
INTERFACE IREADACTIVEALARMSSERVICEPROVIDER
END_INTERFACE

METHOD GETPROXYACTIVEALARMOBJECT : IProxyAlarmObject
VAR_INPUT
	DIOBJNUM : DINT;
END_VAR
END_METHOD

(* ---- IREMOTEDEVICETRAVERSALCONSUMER.itf ---- *)
INTERFACE IREMOTEDEVICETRAVERSALCONSUMER
END_INTERFACE

METHOD REMOTEDEVICEREACHED
VAR_INPUT
	ROW : REFERENCE TO AlarmStorageRow;
	XFIRST : BOOL;
	IVERSION : INT;
END_VAR
END_METHOD

(* ---- IRESETVALUEPROVIDER.itf ---- *)
INTERFACE IRESETVALUEPROVIDER
END_INTERFACE

METHOD RESETVALUE : BOOL
VAR_INPUT
	UIID : ALARM_ID;
END_VAR
END_METHOD

(* ---- ISERVICECONSUMER.itf ---- *)
INTERFACE ISERVICECONSUMER
END_INTERFACE

METHOD ERRORADDED
VAR_INPUT
	UDIERROR : UDINT;
	SMSG : STRING;
	STASKNAME : STRING;
END_VAR
END_METHOD

METHOD REQUESTCLOSED
VAR_INPUT
	IREQUESTID : INT;
END_VAR
END_METHOD

METHOD SETERRORFROMDEVICE
VAR_INPUT
	IERROR : INT;
END_VAR
END_METHOD

(* ---- ISERVICEPROVIDER.itf ---- *)
INTERFACE ISERVICEPROVIDER
END_INTERFACE

METHOD GETAPPLICATION : STRING
END_METHOD

METHOD GETDEVICENAME : STRING
END_METHOD

METHOD GETRECORDID : INT
END_METHOD

(* ---- ISTUBSERVICEMETAOBJECT.itf ---- *)
INTERFACE ISTUBSERVICEMETAOBJECT
END_INTERFACE

METHOD FILLINGCOMPLETED : UDINT
END_METHOD

(* ---- ITAGGEDSERVICEWRITER.itf ---- *)
INTERFACE ITAGGEDSERVICEWRITER
END_INTERFACE

METHOD WRITEBYTE : UDINT
VAR_INPUT
	BT : BYTE;
END_VAR
END_METHOD

METHOD WRITECOMPLEXSTARTTAG : UDINT
VAR_INPUT
	UDITAG : UDINT;
	UDIMINLENSIZE : UDINT;
END_VAR
END_METHOD

METHOD WRITEDWORD : UDINT
VAR_INPUT
	DW : DWORD;
END_VAR
END_METHOD

METHOD WRITEDATASTARTTAG : UDINT
VAR_INPUT
	UDITAG : UDINT;
	ALIGNMENT : CmpBinTagUtilIec.BTagAlignment;
	UDIMINLENSIZE : UDINT;
END_VAR
END_METHOD

METHOD WRITEENDTAG : UDINT
VAR_INPUT
	UDITAG : UDINT;
END_VAR
END_METHOD

METHOD WRITEFILLBYTES : UDINT
END_METHOD

METHOD WRITELWORD : UDINT
VAR_INPUT
	LW : LWORD;
END_VAR
END_METHOD

METHOD WRITESTRING : UDINT
VAR_INPUT
	PSSTRING : POINTER TO STRING(255);
END_VAR
END_METHOD

METHOD WRITEWSTRING : UDINT
VAR_INPUT
	PWSSTRING : POINTER TO WSTRING(255);
END_VAR
END_METHOD

METHOD WRITEWORD : UDINT
VAR_INPUT
	WD : WORD;
END_VAR
END_METHOD

(* ---- IVALUEPROVIDER.itf ---- *)
INTERFACE IVALUEPROVIDER
END_INTERFACE

METHOD GETVALUE : __SYSTEM.TYPE_CLASS
VAR_INPUT
	UIID : ALARM_ID;
	EWHICHVALUE : ConfigurableExpression;
	PBYBUFFER : POINTER TO BYTE;
	IBUFFERSIZE : INT;
END_VAR
END_METHOD

(* ---- _GETALARMSFROMSTORAGE.pou ---- *)
FUNCTION _GETALARMSFROMSTORAGE : BOOL
VAR_INPUT
	ISKIPROWS : INT;
	IMAXROWS : INT;
	PSTARRALARMGROUPS : POINTER TO ARRAY [0..0] OF UDINT;
	ICOUNTALARMGROUPS : INT;
	BALLALARMGROUPS : BOOL;
	PSTARRALARMCLASSES : POINTER TO ARRAY [0..0] OF UDINT;
	ICOUNTALARMCLASSES : INT;
	BALLALARMCLASSES : BOOL;
	USIPRIORITYFROM : USINT;
	USIPRIORITYTO : USINT;
	ALARMDATABLOCK : IAlarmDataBlockBase2;
END_VAR
VAR_IN_OUT
	BROWIDVALID : BOOL;
	DIROWID : DINT;
END_VAR
END_FUNCTION

(* ---- _GETCOUNTALARMSFROMSTORAGE.pou ---- *)
FUNCTION _GETCOUNTALARMSFROMSTORAGE : DINT
VAR_INPUT
	PSTARRALARMGROUPS : POINTER TO ARRAY [0..0] OF UDINT;
	ICOUNTALARMGROUPS : INT;
	BALLALARMGROUPS : BOOL;
	PSTARRALARMCLASSES : POINTER TO ARRAY [0..0] OF UDINT;
	ICOUNTALARMCLASSES : INT;
	BALLALARMCLASSES : BOOL;
	USIPRIORITYFROM : USINT;
	USIPRIORITYTO : USINT;
	ALARMDATABLOCK : IAlarmDataBlockBase2;
END_VAR
END_FUNCTION

(* ---- _GETCURRENTROW.pou ---- *)
FUNCTION _GETCURRENTROW : STO.IRow
VAR_INPUT
	ITFCURSOR : STO.ICursor;
END_VAR
VAR_OUTPUT
	EERROR : STO.ERROR;
END_VAR
END_FUNCTION

(* ---- _GETMINMAXROWIDS.pou ---- *)
FUNCTION _GETMINMAXROWIDS : BOOL
VAR_INPUT
	ITFTABLE : STO.ITable;
END_VAR
VAR_OUTPUT
	IDROWMIN : LINT;
	IDROWMAX : LINT;
	EERROR : STO.ERROR;
END_VAR
END_FUNCTION

(* ---- _GETNUMOFROWS.pou ---- *)
FUNCTION _GETNUMOFROWS : CAA.COUNT
VAR_INPUT
	ITFTABLE : STO.ITable;
END_VAR
VAR_OUTPUT
	EERROR : STO.ERROR;
END_VAR
END_FUNCTION

(* ---- _OPENCURSOR.pou ---- *)
FUNCTION _OPENCURSOR : STO.ICursor
VAR_INPUT
	ITFTABLE : STO.ITable;
	IDINDEX : CAA.IDENT;
	ICOUNTRETRIES : INT;
END_VAR
VAR_OUTPUT
	EERROR : STO.ERROR;
END_VAR
END_FUNCTION

(* ---- ALARMFCTGETLOCALBYTEORDER.pou ---- *)
FUNCTION ALARMFCTGETLOCALBYTEORDER : EAlarmByteOrder
END_FUNCTION
